// TIA Portal V20 program export: 0 tag tables, 60 data types, 15 data blocks, 199 code blocks (in call order from the OBs), 5 instance data blocks

TYPE "FRK_Access"
// stored: IsFailsafeCompliant false
   STRUCT
      CurrentLevel : DInt;
      CurrentUser : String[32];
      LoginFailed : Bool;
      Policy { S7_SetPoint := 'True'} : "ST_AccessPolicy";
      SessionGeneration : UDInt;
      LoginBusy : Bool;
      LoginResultSequence : UDInt;
      LoginTimeoutMs : UDInt;
      PolicySlot { ExternalAccessible := 'False'; ExternalVisible := 'False'; ExternalWritable := 'False'} : Int;
      PolicyLost { ExternalAccessible := 'False'; ExternalVisible := 'False'; ExternalWritable := 'False'} : Bool;
      PolicyLossAlarm { ExternalAccessible := 'False'; ExternalVisible := 'False'; ExternalWritable := 'False'} : Int;
      UserLossAlarm { ExternalAccessible := 'False'; ExternalVisible := 'False'; ExternalWritable := 'False'} : Int;
      ProviderGeneration { ExternalAccessible := 'False'; ExternalVisible := 'False'; ExternalWritable := 'False'} : UDInt;
      CandidateGeneration { ExternalAccessible := 'False'; ExternalVisible := 'False'; ExternalWritable := 'False'} : UDInt;
      ProviderEnabled { ExternalAccessible := 'False'; ExternalVisible := 'False'; ExternalWritable := 'False'} : Bool;
      LastActivity { ExternalAccessible := 'False'; ExternalVisible := 'False'; ExternalWritable := 'False'} : UDInt;
      LoginSince { ExternalAccessible := 'False'; ExternalVisible := 'False'; ExternalWritable := 'False'} : UDInt;
      LoginSequence { ExternalAccessible := 'False'; ExternalVisible := 'False'; ExternalWritable := 'False'} : UDInt;
      CandidateUser { ExternalAccessible := 'False'; ExternalVisible := 'False'; ExternalWritable := 'False'} : String[32];
      CandidateLevel { ExternalAccessible := 'False'; ExternalVisible := 'False'; ExternalWritable := 'False'} : DInt;
      Round { ExternalAccessible := 'False'; ExternalVisible := 'False'; ExternalWritable := 'False'} : DInt;
      Salt { ExternalAccessible := 'False'; ExternalVisible := 'False'; ExternalWritable := 'False'} : Array[0..15] of Byte;
      Digest { ExternalAccessible := 'False'; ExternalVisible := 'False'; ExternalWritable := 'False'} : Array[0..31] of Byte;
      Expected { ExternalAccessible := 'False'; ExternalVisible := 'False'; ExternalWritable := 'False'} : Array[0..31] of Byte;
   END_STRUCT;
END_TYPE

TYPE "FRK_AccessPolicyImage"
// stored: IsFailsafeCompliant false
   STRUCT
      SchemaVersion { ExternalAccessible := 'False'; ExternalVisible := 'False'; ExternalWritable := 'False'} : UInt;
      Initialized { ExternalAccessible := 'False'; ExternalVisible := 'False'; ExternalWritable := 'False'} : Bool;
      Scope { ExternalAccessible := 'False'; ExternalVisible := 'False'; ExternalWritable := 'False'} : String[80];
      Generation { ExternalAccessible := 'False'; ExternalVisible := 'False'; ExternalWritable := 'False'} : UDInt;
      Policy { ExternalAccessible := 'False'; ExternalVisible := 'False'; ExternalWritable := 'False'; S7_SetPoint := 'True'} : "ST_AccessPolicy";
      Checksum { ExternalAccessible := 'False'; ExternalVisible := 'False'; ExternalWritable := 'False'} : DWord;
   END_STRUCT;
END_TYPE

TYPE "FRK_AlarmLog"
// stored: IsFailsafeCompliant false
   STRUCT
      Active { S7_SetPoint := 'True'} : Array[1..16] of "ST_AlarmEvent";
      NActive : Int;
      Ring { S7_SetPoint := 'True'} : Array[1..64] of "ST_AlarmEvent";
      RingHead : Int;
      Blocking : Bool;
      Truncated : Bool;
      ComeMs { ExternalAccessible := 'False'; ExternalVisible := 'False'; ExternalWritable := 'False'} : Array[1..16] of UDInt;
      Automatic { ExternalAccessible := 'False'; ExternalVisible := 'False'; ExternalWritable := 'False'} : Array[1..16] of Bool;
      Touched { ExternalAccessible := 'False'; ExternalVisible := 'False'; ExternalWritable := 'False'} : Array[1..16] of Bool;
      RingUsed { ExternalAccessible := 'False'; ExternalVisible := 'False'; ExternalWritable := 'False'} : Int;
   END_STRUCT;
END_TYPE

TYPE "FRK_Carrier"
// stored: IsFailsafeCompliant false
   STRUCT
      Enabled { ExternalAccessible := 'False'; ExternalVisible := 'False'; ExternalWritable := 'False'} : Bool;
      Kind { ExternalAccessible := 'False'; ExternalVisible := 'False'; ExternalWritable := 'False'} : DInt;
      Serial { ExternalAccessible := 'False'; ExternalVisible := 'False'; ExternalWritable := 'False'} : UDInt;
      Context { ExternalAccessible := 'False'; ExternalVisible := 'False'; ExternalWritable := 'False'; S7_SetPoint := 'True'} : "ST_PartContext";
      Written { ExternalAccessible := 'False'; ExternalVisible := 'False'; ExternalWritable := 'False'; S7_SetPoint := 'True'} : "ST_PartContext";
      Writes { ExternalAccessible := 'False'; ExternalVisible := 'False'; ExternalWritable := 'False'} : UDInt;
   END_STRUCT;
END_TYPE

TYPE "FRK_ConfigCursor"
// stored: IsFailsafeCompliant false
   STRUCT
      Position { ExternalAccessible := 'False'; ExternalVisible := 'False'; ExternalWritable := 'False'} : DInt;
      First { ExternalAccessible := 'False'; ExternalVisible := 'False'; ExternalWritable := 'False'} : DInt;
   END_STRUCT;
END_TYPE

TYPE "FRK_ConfigSlot"
// stored: IsFailsafeCompliant false
   STRUCT
      SchemaVersion { ExternalAccessible := 'False'; ExternalVisible := 'False'; ExternalWritable := 'False'} : UInt;
      Used { ExternalAccessible := 'False'; ExternalVisible := 'False'; ExternalWritable := 'False'} : Bool;
      ModelCode { ExternalAccessible := 'False'; ExternalVisible := 'False'; ExternalWritable := 'False'} : String[64];
      Record { ExternalAccessible := 'False'; ExternalVisible := 'False'; ExternalWritable := 'False'; S7_SetPoint := 'True'} : "ST_ConfigRecord";
   END_STRUCT;
END_TYPE

TYPE "FRK_ConfigValue"
// stored: IsFailsafeCompliant false
   STRUCT
      Number { ExternalAccessible := 'False'; ExternalVisible := 'False'; ExternalWritable := 'False'} : LInt;
      Flag { ExternalAccessible := 'False'; ExternalVisible := 'False'; ExternalWritable := 'False'} : Bool;
      Text { ExternalAccessible := 'False'; ExternalVisible := 'False'; ExternalWritable := 'False'} : String[80];
   END_STRUCT;
END_TYPE

TYPE "FRK_Core"
// stored: IsFailsafeCompliant false
   STRUCT
      Named { ExternalAccessible := 'False'; ExternalVisible := 'False'; ExternalWritable := 'False'} : Bool;
      Initialized { ExternalAccessible := 'False'; ExternalVisible := 'False'; ExternalWritable := 'False'} : Bool;
      RegIndex { ExternalAccessible := 'False'; ExternalVisible := 'False'; ExternalWritable := 'False'} : DInt;
      ParentIndex { ExternalAccessible := 'False'; ExternalVisible := 'False'; ExternalWritable := 'False'} : DInt;
      ModuleType { ExternalAccessible := 'False'; ExternalVisible := 'False'; ExternalWritable := 'False'} : DInt;
      Exec { ExternalAccessible := 'False'; ExternalVisible := 'False'; ExternalWritable := 'False'} : DInt;
      ExecPrev { ExternalAccessible := 'False'; ExternalVisible := 'False'; ExternalWritable := 'False'} : Bool;
      AbortPrev { ExternalAccessible := 'False'; ExternalVisible := 'False'; ExternalWritable := 'False'} : Bool;
      Armed { ExternalAccessible := 'False'; ExternalVisible := 'False'; ExternalWritable := 'False'} : Bool;
      Command { ExternalAccessible := 'False'; ExternalVisible := 'False'; ExternalWritable := 'False'} : DInt;
      CommandLabel { ExternalAccessible := 'False'; ExternalVisible := 'False'; ExternalWritable := 'False'} : String[120];
      Dispatch { ExternalAccessible := 'False'; ExternalVisible := 'False'; ExternalWritable := 'False'} : Bool;
      EvInit { ExternalAccessible := 'False'; ExternalVisible := 'False'; ExternalWritable := 'False'} : Bool;
      EvCommandStart { ExternalAccessible := 'False'; ExternalVisible := 'False'; ExternalWritable := 'False'} : Bool;
      ReleasePending { ExternalAccessible := 'False'; ExternalVisible := 'False'; ExternalWritable := 'False'} : Bool;
      EvAbort { ExternalAccessible := 'False'; ExternalVisible := 'False'; ExternalWritable := 'False'} : Bool;
      EvAbortInError { ExternalAccessible := 'False'; ExternalVisible := 'False'; ExternalWritable := 'False'} : Bool;
      EvModeExit { ExternalAccessible := 'False'; ExternalVisible := 'False'; ExternalWritable := 'False'} : Bool;
      EvModeChanged { ExternalAccessible := 'False'; ExternalVisible := 'False'; ExternalWritable := 'False'} : Bool;
      "Step" { ExternalAccessible := 'False'; ExternalVisible := 'False'; ExternalWritable := 'False'} : DInt;
      HookResult { ExternalAccessible := 'False'; ExternalVisible := 'False'; ExternalWritable := 'False'} : DInt;
      Held { ExternalAccessible := 'False'; ExternalVisible := 'False'; ExternalWritable := 'False'} : Bool;
      HoldReq { ExternalAccessible := 'False'; ExternalVisible := 'False'; ExternalWritable := 'False'} : Bool;
      HoldReason { ExternalAccessible := 'False'; ExternalVisible := 'False'; ExternalWritable := 'False'} : DInt;
      DiagTouched { ExternalAccessible := 'False'; ExternalVisible := 'False'; ExternalWritable := 'False'} : Bool;
      TimingOpen { ExternalAccessible := 'False'; ExternalVisible := 'False'; ExternalWritable := 'False'} : Bool;
      StartMs { ExternalAccessible := 'False'; ExternalVisible := 'False'; ExternalWritable := 'False'} : UDInt;
      LastNowMs { ExternalAccessible := 'False'; ExternalVisible := 'False'; ExternalWritable := 'False'} : UDInt;
      DeltaMs { ExternalAccessible := 'False'; ExternalVisible := 'False'; ExternalWritable := 'False'} : UDInt;
      ActiveMs { ExternalAccessible := 'False'; ExternalVisible := 'False'; ExternalWritable := 'False'} : UDInt;
      TimeoutMs { ExternalAccessible := 'False'; ExternalVisible := 'False'; ExternalWritable := 'False'} : UDInt;
      Timing { ExternalAccessible := 'False'; ExternalVisible := 'False'; ExternalWritable := 'False'; S7_SetPoint := 'True'} : "ST_ModuleTiming";
      FaultSlot { ExternalAccessible := 'False'; ExternalVisible := 'False'; ExternalWritable := 'False'} : Int;
      FaultHandled { ExternalAccessible := 'False'; ExternalVisible := 'False'; ExternalWritable := 'False'} : Bool;
   END_STRUCT;
END_TYPE

TYPE "FRK_DecisionSlot"
// stored: IsFailsafeCompliant false
   STRUCT
      RootIndex { ExternalAccessible := 'False'; ExternalVisible := 'False'; ExternalWritable := 'False'} : DInt;
      Owner { ExternalAccessible := 'False'; ExternalVisible := 'False'; ExternalWritable := 'False'} : DInt;
      Request { ExternalAccessible := 'False'; ExternalVisible := 'False'; ExternalWritable := 'False'; S7_SetPoint := 'True'} : "ST_DecisionRequest";
      Answer { ExternalAccessible := 'False'; ExternalVisible := 'False'; ExternalWritable := 'False'} : Int;
      AskedAt { ExternalAccessible := 'False'; ExternalVisible := 'False'; ExternalWritable := 'False'} : UDInt;
      OverlapLogged { ExternalAccessible := 'False'; ExternalVisible := 'False'; ExternalWritable := 'False'} : Bool;
      ResolutionLogged { ExternalAccessible := 'False'; ExternalVisible := 'False'; ExternalWritable := 'False'} : Bool;
   END_STRUCT;
END_TYPE

TYPE "FRK_JsonField"
// stored: IsFailsafeCompliant false
   STRUCT
      Key { ExternalAccessible := 'False'; ExternalVisible := 'False'; ExternalWritable := 'False'} : String[16];
      Text { ExternalAccessible := 'False'; ExternalVisible := 'False'; ExternalWritable := 'False'} : WString[160];
      Quoted { ExternalAccessible := 'False'; ExternalVisible := 'False'; ExternalWritable := 'False'} : Bool;
   END_STRUCT;
END_TYPE

TYPE "FRK_ManualConditionRow"
// stored: IsFailsafeCompliant false
   STRUCT
      Used { ExternalAccessible := 'False'; ExternalVisible := 'False'; ExternalWritable := 'False'} : Bool;
      Value { ExternalAccessible := 'False'; ExternalVisible := 'False'; ExternalWritable := 'False'} : DInt;
      Ok { ExternalAccessible := 'False'; ExternalVisible := 'False'; ExternalWritable := 'False'} : Bool;
      Diag { ExternalAccessible := 'False'; ExternalVisible := 'False'; ExternalWritable := 'False'; S7_SetPoint := 'True'} : "ST_Diagnostic";
      Bypassable { ExternalAccessible := 'False'; ExternalVisible := 'False'; ExternalWritable := 'False'} : Bool;
   END_STRUCT;
END_TYPE

TYPE "FRK_PermCtx"
// stored: IsFailsafeCompliant false
   STRUCT
      Permit : Bool;
      Count : Int;
      Blocker : String[160];
   END_STRUCT;
END_TYPE

TYPE "FRK_RegistryRow"
// stored: IsFailsafeCompliant false
   STRUCT
      Valid { ExternalAccessible := 'False'; ExternalVisible := 'False'; ExternalWritable := 'False'} : Bool;
      Parent { ExternalAccessible := 'False'; ExternalVisible := 'False'; ExternalWritable := 'False'} : DInt;
      ModuleType { ExternalAccessible := 'False'; ExternalVisible := 'False'; ExternalWritable := 'False'} : DInt;
      TypeId { ExternalAccessible := 'False'; ExternalVisible := 'False'; ExternalWritable := 'False'} : DInt;
      Capabilities { ExternalAccessible := 'False'; ExternalVisible := 'False'; ExternalWritable := 'False'} : DWord;
      Exec { ExternalAccessible := 'False'; ExternalVisible := 'False'; ExternalWritable := 'False'} : DInt;
      ReasonCode { ExternalAccessible := 'False'; ExternalVisible := 'False'; ExternalWritable := 'False'} : DInt;
      Severity { ExternalAccessible := 'False'; ExternalVisible := 'False'; ExternalWritable := 'False'} : DInt;
      AlarmBlocking { ExternalAccessible := 'False'; ExternalVisible := 'False'; ExternalWritable := 'False'} : Bool;
   END_STRUCT;
END_TYPE

TYPE "FRK_SequenceCtx"
// stored: IsFailsafeCompliant false
   STRUCT
      RunPrevious { ExternalAccessible := 'False'; ExternalVisible := 'False'; ExternalWritable := 'False'} : Bool;
      Running : Bool;
      Restart { ExternalAccessible := 'False'; ExternalVisible := 'False'; ExternalWritable := 'False'} : Bool;
      Done : Bool;
      Error : Bool;
      Pending : Bool;
      StartLatched { ExternalAccessible := 'False'; ExternalVisible := 'False'; ExternalWritable := 'False'} : Bool;
      OwnerIndex { ExternalAccessible := 'False'; ExternalVisible := 'False'; ExternalWritable := 'False'} : DInt;
      ChainIndex { ExternalAccessible := 'False'; ExternalVisible := 'False'; ExternalWritable := 'False'} : DInt;
      "Step" : DInt;
      ScanStep { ExternalAccessible := 'False'; ExternalVisible := 'False'; ExternalWritable := 'False'} : DInt;
      RecordedStep { ExternalAccessible := 'False'; ExternalVisible := 'False'; ExternalWritable := 'False'} : DInt;
      RetVal { ExternalAccessible := 'False'; ExternalVisible := 'False'; ExternalWritable := 'False'} : DInt;
      Scan { ExternalAccessible := 'False'; ExternalVisible := 'False'; ExternalWritable := 'False'} : UDInt;
      Visit { ExternalAccessible := 'False'; ExternalVisible := 'False'; ExternalWritable := 'False'} : UDInt;
      Elapsed : Time;
      DelayElapsed { ExternalAccessible := 'False'; ExternalVisible := 'False'; ExternalWritable := 'False'} : Time;
      StepName : String[160];
      Awaiting : String[160];
      ErrorDiagnostic { S7_SetPoint := 'True'} : "ST_Diagnostic";
      BranchIndex { ExternalAccessible := 'False'; ExternalVisible := 'False'; ExternalWritable := 'False'} : DInt;
      CommandFailed { ExternalAccessible := 'False'; ExternalVisible := 'False'; ExternalWritable := 'False'} : Bool;
      CommandIssued { ExternalAccessible := 'False'; ExternalVisible := 'False'; ExternalWritable := 'False'} : Bool;
      Warned { ExternalAccessible := 'False'; ExternalVisible := 'False'; ExternalWritable := 'False'} : Bool;
      HandledDiagnostic { ExternalAccessible := 'False'; ExternalVisible := 'False'; ExternalWritable := 'False'; S7_SetPoint := 'True'} : "ST_Diagnostic";
      EventVisit { ExternalAccessible := 'False'; ExternalVisible := 'False'; ExternalWritable := 'False'} : UDInt;
      EventToken { ExternalAccessible := 'False'; ExternalVisible := 'False'; ExternalWritable := 'False'} : DInt;
   END_STRUCT;
END_TYPE

TYPE "FRK_SequenceRow"
// stored: IsFailsafeCompliant false
   STRUCT
      StepNo : DInt;
      Visited : Bool;
      LastDuration : Time;
   END_STRUCT;
END_TYPE

TYPE "FRK_SetPayload"
// stored: IsFailsafeCompliant false
   STRUCT
      Info { ExternalAccessible := 'False'; ExternalVisible := 'False'; ExternalWritable := 'False'; S7_SetPoint := 'True'} : "ST_ConfigSetInfo";
      Records { ExternalAccessible := 'False'; ExternalVisible := 'False'; ExternalWritable := 'False'; S7_SetPoint := 'True'} : Array[1..3] of "ST_ConfigRecord";
   END_STRUCT;
END_TYPE

TYPE "FRK_SetWorkspace"
// stored: IsFailsafeCompliant false
   STRUCT
      Payload { ExternalAccessible := 'False'; ExternalVisible := 'False'; ExternalWritable := 'False'; S7_SetPoint := 'True'} : "FRK_SetPayload";
      Seen { ExternalAccessible := 'False'; ExternalVisible := 'False'; ExternalWritable := 'False'} : Array[1..3] of Bool;
      Matched { ExternalAccessible := 'False'; ExternalVisible := 'False'; ExternalWritable := 'False'} : Int;
      RejectScope { ExternalAccessible := 'False'; ExternalVisible := 'False'; ExternalWritable := 'False'} : String[80];
      RejectKey { ExternalAccessible := 'False'; ExternalVisible := 'False'; ExternalWritable := 'False'} : String[160];
      Importing { ExternalAccessible := 'False'; ExternalVisible := 'False'; ExternalWritable := 'False'} : Bool;
      Exporting { ExternalAccessible := 'False'; ExternalVisible := 'False'; ExternalWritable := 'False'} : Bool;
      NextLine { ExternalAccessible := 'False'; ExternalVisible := 'False'; ExternalWritable := 'False'} : Int;
      Generation { ExternalAccessible := 'False'; ExternalVisible := 'False'; ExternalWritable := 'False'} : UDInt;
      Received { ExternalAccessible := 'False'; ExternalVisible := 'False'; ExternalWritable := 'False'} : Int;
      Piece { ExternalAccessible := 'False'; ExternalVisible := 'False'; ExternalWritable := 'False'} : WString[480];
      Line { ExternalAccessible := 'False'; ExternalVisible := 'False'; ExternalWritable := 'False'} : WString[480];
      Fields { ExternalAccessible := 'False'; ExternalVisible := 'False'; ExternalWritable := 'False'; S7_SetPoint := 'True'} : Array[1..9] of "FRK_JsonField";
      FieldCount { ExternalAccessible := 'False'; ExternalVisible := 'False'; ExternalWritable := 'False'} : Int;
   END_STRUCT;
END_TYPE

TYPE "FRK_Unit"
// stored: IsFailsafeCompliant false
   STRUCT
      Initialized { ExternalAccessible := 'False'; ExternalVisible := 'False'; ExternalWritable := 'False'} : Bool;
      Mode { ExternalAccessible := 'False'; ExternalVisible := 'False'; ExternalWritable := 'False'} : DInt;
      RequestedMode { ExternalAccessible := 'False'; ExternalVisible := 'False'; ExternalWritable := 'False'} : DInt;
      ModePending { ExternalAccessible := 'False'; ExternalVisible := 'False'; ExternalWritable := 'False'} : Bool;
      ExitFirst { ExternalAccessible := 'False'; ExternalVisible := 'False'; ExternalWritable := 'False'} : Bool;
      RunReq { ExternalAccessible := 'False'; ExternalVisible := 'False'; ExternalWritable := 'False'} : Bool;
      AbortReq { ExternalAccessible := 'False'; ExternalVisible := 'False'; ExternalWritable := 'False'} : Bool;
      StopReq { ExternalAccessible := 'False'; ExternalVisible := 'False'; ExternalWritable := 'False'} : Bool;
      ModeSince { ExternalAccessible := 'False'; ExternalVisible := 'False'; ExternalWritable := 'False'} : UDInt;
      ReleaseChildren { ExternalAccessible := 'False'; ExternalVisible := 'False'; ExternalWritable := 'False'} : Bool;
      Clearing { ExternalAccessible := 'False'; ExternalVisible := 'False'; ExternalWritable := 'False'} : Bool;
      FaultLatched { ExternalAccessible := 'False'; ExternalVisible := 'False'; ExternalWritable := 'False'} : Bool;
      PrevError { ExternalAccessible := 'False'; ExternalVisible := 'False'; ExternalWritable := 'False'} : Bool;
      EvReset { ExternalAccessible := 'False'; ExternalVisible := 'False'; ExternalWritable := 'False'} : Bool;
      SeenSequence { ExternalAccessible := 'False'; ExternalVisible := 'False'; ExternalWritable := 'False'} : UDInt;
      RequestPending { ExternalAccessible := 'False'; ExternalVisible := 'False'; ExternalWritable := 'False'} : Bool;
      Request { ExternalAccessible := 'False'; ExternalVisible := 'False'; ExternalWritable := 'False'; S7_SetPoint := 'True'} : "ST_HmiRequest";
      RequestUser { ExternalAccessible := 'False'; ExternalVisible := 'False'; ExternalWritable := 'False'} : String[32];
      Permit { ExternalAccessible := 'False'; ExternalVisible := 'False'; ExternalWritable := 'False'} : Bool;
      PermitDiag { ExternalAccessible := 'False'; ExternalVisible := 'False'; ExternalWritable := 'False'; S7_SetPoint := 'True'} : "ST_Diagnostic";
      CarrierIndex { ExternalAccessible := 'False'; ExternalVisible := 'False'; ExternalWritable := 'False'} : DInt;
      Good { ExternalAccessible := 'False'; ExternalVisible := 'False'; ExternalWritable := 'False'} : UDInt;
      Nok { ExternalAccessible := 'False'; ExternalVisible := 'False'; ExternalWritable := 'False'} : UDInt;
      Rework { ExternalAccessible := 'False'; ExternalVisible := 'False'; ExternalWritable := 'False'} : UDInt;
      NokReason { ExternalAccessible := 'False'; ExternalVisible := 'False'; ExternalWritable := 'False'} : DInt;
      CascadePending { ExternalAccessible := 'False'; ExternalVisible := 'False'; ExternalWritable := 'False'} : Bool;
      CascadeKind { ExternalAccessible := 'False'; ExternalVisible := 'False'; ExternalWritable := 'False'} : DInt;
      CascadeMode { ExternalAccessible := 'False'; ExternalVisible := 'False'; ExternalWritable := 'False'} : DInt;
      FollowStart { ExternalAccessible := 'False'; ExternalVisible := 'False'; ExternalWritable := 'False'} : Bool;
      AlarmBlocking { ExternalAccessible := 'False'; ExternalVisible := 'False'; ExternalWritable := 'False'} : Bool;
      ConfigBlocked { ExternalAccessible := 'False'; ExternalVisible := 'False'; ExternalWritable := 'False'} : Bool;
      ConfigEnabled { ExternalAccessible := 'False'; ExternalVisible := 'False'; ExternalWritable := 'False'} : Bool;
      ModelEnabled { ExternalAccessible := 'False'; ExternalVisible := 'False'; ExternalWritable := 'False'} : Bool;
      ConfigSetsEnabled { ExternalAccessible := 'False'; ExternalVisible := 'False'; ExternalWritable := 'False'} : Bool;
   END_STRUCT;
END_TYPE

TYPE "ST_AccessPolicy"
// stored: IsFailsafeCompliant false
   STRUCT
      Required : Array[0..11] of DInt;
      SessionTimeout : Time := T#0MS;
   END_STRUCT;
END_TYPE

TYPE "ST_AlarmEvent"
// stored: IsFailsafeCompliant false
   STRUCT
      ReasonCode : DInt;
      Description : WString[255];
      SourcePath : WString[255];
      IoTag : String[80];
      IoAddress : String[80];
      Severity : DInt;
      Category : DInt;
      ResetClass : DInt;
      State : DInt;
      ComeAt : LDT;
      GoneAt : LDT;
      ResetAt : LDT;
      Duration : Time;
      Shelved : Bool;
      ShelvedUntil : LDT;
      ComeTimeSynchronized : Bool;
      GoneTimeSynchronized : Bool;
      ResetTimeSynchronized : Bool;
      ShelfTimeSynchronized : Bool;
   END_STRUCT;
END_TYPE

TYPE "ST_CommandInfo"
// stored: IsFailsafeCompliant false
   STRUCT
      Value : DInt;
      Label : String[120];
      Style : DInt;
   END_STRUCT;
END_TYPE

TYPE "ST_ConfigEntry"
// stored: IsFailsafeCompliant false
   STRUCT
      Scope : WString[255];
      Item : WString[255];
      ValueText : WString[255];
      WriteKey : String[160];
      WriteRevision : UDInt;
      ConfigKind : DInt;
      ValueType : DInt;
      Writable : Bool;
      RequiresReady : Bool;
      HasMinimum : Bool;
      HasMaximum : Bool;
      Minimum : LReal;
      Maximum : LReal;
      Unit : String[16];
      LabelKey : String[160];
      EnumDomain : WString[255];
      ClassId : String[40];
      ReadLevel : DInt;
      WriteLevel : DInt;
      Readable : Bool;
      UnitCode : DInt;
      EnumLabelKey : String[80];
      ModelScoped : Bool;
   END_STRUCT;
END_TYPE

TYPE "ST_ConfigPage"
// stored: IsFailsafeCompliant false
   STRUCT
      Revision : UDInt;
      PageIndex : Int;
      PageCount : Int;
      EntryCount : Int;
      Entries { S7_SetPoint := 'True'} : Array[1..16] of "ST_ConfigEntry";
   END_STRUCT;
END_TYPE

TYPE "ST_ConfigPersistStatus"
// stored: IsFailsafeCompliant false
   STRUCT
      Pending : Bool;
      Failed : Bool;
      WindowMs : UDInt := 5000;
      PendingSince : LDT;
      StorePresent : Bool;
      StoreKind : DInt;
      RestorePolicy : DInt;
      RestoreLost : Bool;
      RestoreAcknowledged : Bool;
      LostPath : String[80];
      LastSetName : String[80];
      LastSetRecords : Int;
      LastRejectScope : String[80];
      LastRejectKey : String[160];
   END_STRUCT;
END_TYPE

TYPE "ST_ConfigRecord"
// stored: IsFailsafeCompliant false
   STRUCT
      Scope : String[80];
      WriteKey : String[160];
      Revision : UDInt;
      Kind : DInt;
      ValueType : DInt;
      ValueText : String[80];
   END_STRUCT;
END_TYPE

TYPE "ST_ConfigSetInfo"
// stored: IsFailsafeCompliant false
   STRUCT
      Used : Bool;
      SetName : String[80];
      RootIdentity : String[80];
      SetSchema : UInt;
      ConfigRev : UDInt;
      Kind : DInt;
      ModelCode : String[64];
      RecordCount : Int;
      CreatedAt : LDT;
      TimeSynchronized : Bool;
   END_STRUCT;
END_TYPE

TYPE "ST_CylinderDevice"
// stored: IsFailsafeCompliant false
   STRUCT
      Direction : DInt;
      Withdrawn : Bool;
      Extended : Bool;
      Retracted : Bool;
      Lease { S7_SetPoint := 'True'} : "ST_SequenceCommandLease";
   END_STRUCT;
END_TYPE

TYPE "ST_CylinderHal"
// stored: IsFailsafeCompliant false
   STRUCT
      FeedbackExtended : Bool;
      FeedbackRetracted : Bool;
      ExtendPermit : Bool;
      RetractPermit : Bool;
      PermitDiagnostic { S7_SetPoint := 'True'} : "ST_Diagnostic";
      RetractDiagnostic { S7_SetPoint := 'True'} : "ST_Diagnostic";
      CoilExtend : Bool;
      CoilRetract : Bool;
   END_STRUCT;
END_TYPE

TYPE "ST_CylinderOutCmd"
// stored: IsFailsafeCompliant false
   STRUCT
      Direction : DInt;
   END_STRUCT;
END_TYPE

TYPE "ST_CylinderOutImm"
// stored: IsFailsafeCompliant false
   STRUCT
      Extended : Bool;
      Retracted : Bool;
   END_STRUCT;
END_TYPE

TYPE "ST_CylinderParCfg"
// stored: IsFailsafeCompliant false
   STRUCT
      SchemaVersion : UInt := 1;
      Timeout : Time := T#8S;
   END_STRUCT;
END_TYPE

TYPE "ST_CylinderParCmd"
// stored: IsFailsafeCompliant false
   STRUCT
      Reserved : Bool;
   END_STRUCT;
END_TYPE

TYPE "ST_DecisionRequest"
// stored: IsFailsafeCompliant false
   STRUCT
      Prompt : WString[255];
      Options : Array[1..6] of String[64];
      Default : Int;
      Timeout : Time;
      SourcePath : WString[255];
   END_STRUCT;
END_TYPE

TYPE "ST_Diagnostic"
// stored: IsFailsafeCompliant false
   STRUCT
      ReasonCode : DInt;
      SourcePath : WString[255];
      Description : WString[255];
      IoTag : String[80];
      IoAddress : String[80];
      Severity : DInt;
      Category : DInt;
      Since : LDT;
      TimeSynchronized : Bool;
   END_STRUCT;
END_TYPE

TYPE "ST_FraktalHal"
// stored: IsFailsafeCompliant false
   STRUCT
      PressDemo { ExternalAccessible := 'False'; ExternalVisible := 'False'; ExternalWritable := 'False'; S7_SetPoint := 'True'} : "ST_PressDemoUnitHal";
   END_STRUCT;
END_TYPE

TYPE "ST_HmiRequest"
// stored: IsFailsafeCompliant false
   STRUCT
      Kind : DInt;
      TargetPath : WString[255];
      NameValue : String[160];
      TextValue : WString[255];
      User : String[32];
      Secret : String[32];
      IntValue : DInt;
      BoolValue : Bool;
      DurationMs : UDInt;
      Sequence : UDInt;
   END_STRUCT;
END_TYPE

TYPE "ST_HmiResponse"
// stored: IsFailsafeCompliant false
   STRUCT
      AckSequence : UDInt;
      Accepted : Bool;
      Diagnostic : WString[255];
      Report { S7_SetPoint := 'True'} : "ST_ReleaseReport";
      ConfigPage { S7_SetPoint := 'True'} : "ST_ConfigPage";
   END_STRUCT;
END_TYPE

TYPE "ST_MeasRecord"
// stored: IsFailsafeCompliant false
   STRUCT
      "Name" : String[64];
      Value : LReal;
      Minimum : LReal;
      Maximum : LReal;
      Target : LReal;
      Unit : String[16];
      InTol : Bool;
   END_STRUCT;
END_TYPE

TYPE "ST_ModePolicy"
// stored: IsFailsafeCompliant false
   STRUCT
      Shield : DInt;
      Style : DInt;
   END_STRUCT;
END_TYPE

TYPE "ST_ModelField"
// stored: IsFailsafeCompliant false
   STRUCT
      "Name" : String[32];
      Value : String[64];
   END_STRUCT;
END_TYPE

TYPE "ST_ModelId"
// stored: IsFailsafeCompliant false
   STRUCT
      ModelCode : String[64];
      "Family" : String[64];
      Variant : String[64];
      Fields { S7_SetPoint := 'True'} : Array[1..8] of "ST_ModelField";
      NField : Int;
   END_STRUCT;
END_TYPE

TYPE "ST_ModuleStatus"
// stored: IsFailsafeCompliant false
   STRUCT
      "Name" : String[80];
      DisplayNameKey : String[160];
      DescriptionKey : String[160];
      TypeKey : String[160];
      ModuleType : DInt;
      State : DInt;
      FaultActive : Bool;
      Diagnostic { S7_SetPoint := 'True'} : "ST_Diagnostic";
      TileEnable : Bool := TRUE;
      ControlDomainId : String[80];
   END_STRUCT;
END_TYPE

TYPE "ST_ModuleTiming"
// stored: IsFailsafeCompliant false
   STRUCT
      LastCmdTime : Time;
      Rows { S7_SetPoint := 'True'} : Array[1..8] of "ST_TimingRow";
      Truncated : Bool;
   END_STRUCT;
END_TYPE

TYPE "ST_PartContext"
// stored: IsFailsafeCompliant false
   STRUCT
      Uid : String[64];
      Present : Bool;
      CarrierKind : DInt;
      Result { S7_SetPoint := 'True'} : "ST_PartResult";
      Parents : Array[1..8] of String[64];
   END_STRUCT;
END_TYPE

TYPE "ST_PartResult"
// stored: IsFailsafeCompliant false
   STRUCT
      Verdict : DInt;
      ReasonCode : DInt;
      Records { S7_SetPoint := 'True'} : Array[1..32] of "ST_MeasRecord";
      StationPath : WString[255];
      Stamp : LDT;
      TimeSynchronized : Bool;
   END_STRUCT;
END_TYPE

TYPE "ST_PressDemoCycle"
// stored: IsFailsafeCompliant false
   STRUCT
      PartInMachine { ExternalAccessible := 'False'; ExternalVisible := 'False'; ExternalWritable := 'False'} : Bool;
      PartDispositioned { ExternalAccessible := 'False'; ExternalVisible := 'False'; ExternalWritable := 'False'} : Bool;
      CycleCompleted { ExternalAccessible := 'False'; ExternalVisible := 'False'; ExternalWritable := 'False'} : Bool;
      FailureReason { ExternalAccessible := 'False'; ExternalVisible := 'False'; ExternalWritable := 'False'} : DInt;
   END_STRUCT;
END_TYPE

TYPE "ST_PressDemoOutCmd"
// stored: IsFailsafeCompliant false
   STRUCT
      CycleCompleted : Bool;
   END_STRUCT;
END_TYPE

TYPE "ST_PressDemoOutImm"
// stored: IsFailsafeCompliant false
   STRUCT
      Homed : Bool;
   END_STRUCT;
END_TYPE

TYPE "ST_PressDemoParCfg"
// stored: IsFailsafeCompliant false
   STRUCT
      SchemaVersion : UInt := 1;
      Timeout : Time := T#0MS;
   END_STRUCT;
END_TYPE

TYPE "ST_PressDemoParCmd"
// stored: IsFailsafeCompliant false
   STRUCT
      Reserved : Bool;
   END_STRUCT;
END_TYPE

TYPE "ST_PressDemoReleaseConditions"
// stored: IsFailsafeCompliant false
   STRUCT
      ModeStartAirPressureOk : Bool;
      RamGuardClosed : Bool;
      RamSlideInside : Bool;
      RamDevicesHealthy : Bool;
      RamAirPressureOk : Bool;
      RamTwoHandHeld : Bool;
   END_STRUCT;
END_TYPE

TYPE "ST_PressDemoSignals"
// stored: IsFailsafeCompliant false
   STRUCT
      PartPresent { ExternalAccessible := 'False'; ExternalVisible := 'False'; ExternalWritable := 'False'} : Bool;
      PartQuality { ExternalAccessible := 'False'; ExternalVisible := 'False'; ExternalWritable := 'False'} : Bool;
      AirPressureOk { ExternalAccessible := 'False'; ExternalVisible := 'False'; ExternalWritable := 'False'} : Bool;
      TwoHandHeld { ExternalAccessible := 'False'; ExternalVisible := 'False'; ExternalWritable := 'False'} : Bool;
      StartPulse { ExternalAccessible := 'False'; ExternalVisible := 'False'; ExternalWritable := 'False'} : Bool;
      PermitDiagnostic { ExternalAccessible := 'False'; ExternalVisible := 'False'; ExternalWritable := 'False'; S7_SetPoint := 'True'} : "ST_Diagnostic";
   END_STRUCT;
END_TYPE

TYPE "ST_PressDemoStationCfg"
// stored: IsFailsafeCompliant false
   STRUCT
      SchemaVersion : UInt := 1;
      RequireTwoHandStart : Bool := TRUE;
      TransferSettleTime : Time := T#200MS;
      PressSettleTime : Time := T#300MS;
   END_STRUCT;
END_TYPE

TYPE "ST_PressDemoUnitHal"
// stored: IsFailsafeCompliant false
   STRUCT
      PressRam { ExternalAccessible := 'False'; ExternalVisible := 'False'; ExternalWritable := 'False'; S7_SetPoint := 'True'} : "ST_CylinderHal";
      Door { ExternalAccessible := 'False'; ExternalVisible := 'False'; ExternalWritable := 'False'; S7_SetPoint := 'True'} : "ST_CylinderHal";
      PartSlide { ExternalAccessible := 'False'; ExternalVisible := 'False'; ExternalWritable := 'False'; S7_SetPoint := 'True'} : "ST_CylinderHal";
      Process { ExternalAccessible := 'False'; ExternalVisible := 'False'; ExternalWritable := 'False'; S7_SetPoint := 'True'} : "ST_PressDemoSignals";
   END_STRUCT;
END_TYPE

TYPE "ST_ReleaseReason"
// stored: IsFailsafeCompliant false
   STRUCT
      Description : WString[255];
      ReasonCode : DInt;
      SourcePath : WString[255];
      Kind : DInt;
      Bypassable : Bool;
   END_STRUCT;
END_TYPE

TYPE "ST_ReleaseReport"
// stored: IsFailsafeCompliant false
   STRUCT
      Released : Bool;
      Count : Int;
      Reasons { S7_SetPoint := 'True'} : Array[1..24] of "ST_ReleaseReason";
   END_STRUCT;
END_TYPE

TYPE "ST_SequenceCommandLease"
// stored: IsFailsafeCompliant false
   STRUCT
      OwnerIndex : DInt;
      ChainIndex : DInt;
      BranchIndex : DInt;
      "Step" : DInt;
      Raised : Bool;
      AbortIssued : Bool;
      ReleasedScan : UDInt;
   END_STRUCT;
END_TYPE

TYPE "ST_StateFlag"
// stored: IsFailsafeCompliant false
   STRUCT
      Key : String[120];
      Value : Bool;
      Since : LDT;
      Stale : Bool;
   END_STRUCT;
END_TYPE

TYPE "ST_TimingRow"
// stored: IsFailsafeCompliant false
   STRUCT
      Id : DInt;
      Label : String[120];
      TimeClass : DInt;
      Count : UDInt;
      Last : Time;
      Minimum : Time;
      Maximum : Time;
      Avg : Time;
   END_STRUCT;
END_TYPE

TYPE "ST_UserRecord"
// stored: IsFailsafeCompliant false
   STRUCT
      User : String[32];
      Salt : Array[0..15] of Byte;
      PinHash : Array[0..31] of Byte;
      Level : DInt;
   END_STRUCT;
END_TYPE

DATA_BLOCK "FRK_AccessPolicies"   // DB3
{ S7_Optimized_Access := 'TRUE' }
VERSION : 0.1
// stored: AutoNumber true, DBAccessibleFromOPCUA true, DBAccessibleFromWebserver true, IsOnlyStoredInLoadMemory false, IsRetainMemResEnabled false, IsWriteProtectedInAS false, MemoryReserve 100
   VAR RETAIN
      Rows { ExternalAccessible := 'False'; ExternalVisible := 'False'; ExternalWritable := 'False'; S7_SetPoint := 'True'} : Array[1..1] of "FRK_AccessPolicyImage";
   END_VAR
BEGIN
END_DATA_BLOCK

DATA_BLOCK "FRK_AccessStorage"   // DB4
{ S7_Optimized_Access := 'TRUE' }
VERSION : 0.1
// stored: AutoNumber true, DBAccessibleFromOPCUA true, DBAccessibleFromWebserver true, IsOnlyStoredInLoadMemory false, IsRetainMemResEnabled false, IsWriteProtectedInAS false, MemoryReserve 100
   VAR
      UsersReady { ExternalAccessible := 'False'; ExternalVisible := 'False'; ExternalWritable := 'False'} : Bool;
      UsersLost { ExternalAccessible := 'False'; ExternalVisible := 'False'; ExternalWritable := 'False'} : Bool;
      EmptyPolicy { ExternalAccessible := 'False'; ExternalVisible := 'False'; ExternalWritable := 'False'; S7_SetPoint := 'True'} : "ST_AccessPolicy";
   END_VAR
   VAR RETAIN
      UsersCommissioned { ExternalAccessible := 'False'; ExternalVisible := 'False'; ExternalWritable := 'False'} : Bool;
   END_VAR
BEGIN
END_DATA_BLOCK

DATA_BLOCK "FRK_Carriers"   // DB5
{ S7_Optimized_Access := 'TRUE' }
VERSION : 0.1
// stored: AutoNumber true, DBAccessibleFromOPCUA true, DBAccessibleFromWebserver true, IsOnlyStoredInLoadMemory false, IsRetainMemResEnabled false, IsWriteProtectedInAS false, MemoryReserve 100
   VAR
      Slots { ExternalAccessible := 'False'; ExternalVisible := 'False'; ExternalWritable := 'False'; S7_SetPoint := 'True'} : Array[0..4] of "FRK_Carrier";
   END_VAR
BEGIN
END_DATA_BLOCK

DATA_BLOCK "FRK_Clock"   // DB1
{ S7_Optimized_Access := 'TRUE' }
VERSION : 0.1
// stored: AutoNumber true, DBAccessibleFromOPCUA true, DBAccessibleFromWebserver true, IsOnlyStoredInLoadMemory false, IsRetainMemResEnabled false, IsWriteProtectedInAS false, MemoryReserve 100
   VAR
      Mem { ExternalAccessible := 'False'; ExternalVisible := 'False'; ExternalWritable := 'False'} : LReal;
      AccMs { ExternalAccessible := 'False'; ExternalVisible := 'False'; ExternalWritable := 'False'} : LReal;
      NowMs { ExternalAccessible := 'False'; ExternalVisible := 'False'; ExternalWritable := 'False'} : UDInt;
   END_VAR
BEGIN
END_DATA_BLOCK

DATA_BLOCK "FRK_ConfigRuntime"   // DB6
{ S7_Optimized_Access := 'TRUE' }
VERSION : 0.1
// stored: AutoNumber true, DBAccessibleFromOPCUA true, DBAccessibleFromWebserver true, IsOnlyStoredInLoadMemory false, IsRetainMemResEnabled false, IsWriteProtectedInAS false, MemoryReserve 100
   VAR
      Fresh { ExternalAccessible := 'False'; ExternalVisible := 'False'; ExternalWritable := 'False'} : Bool;
      Unavailable { ExternalAccessible := 'False'; ExternalVisible := 'False'; ExternalWritable := 'False'} : Bool;
      Failed { ExternalAccessible := 'False'; ExternalVisible := 'False'; ExternalWritable := 'False'} : Array[1..1] of Bool;
      LossSlot { ExternalAccessible := 'False'; ExternalVisible := 'False'; ExternalWritable := 'False'} : Array[1..1] of Int;
   END_VAR
BEGIN
END_DATA_BLOCK

DATA_BLOCK "FRK_ConfigScratch"   // DB7
{ S7_Optimized_Access := 'TRUE' }
VERSION : 0.1
// stored: AutoNumber true, DBAccessibleFromOPCUA true, DBAccessibleFromWebserver true, IsOnlyStoredInLoadMemory false, IsRetainMemResEnabled false, IsWriteProtectedInAS false, MemoryReserve 100
   VAR
      Entry { ExternalAccessible := 'False'; ExternalVisible := 'False'; ExternalWritable := 'False'; S7_SetPoint := 'True'} : "ST_ConfigEntry";
      Blank { ExternalAccessible := 'False'; ExternalVisible := 'False'; ExternalWritable := 'False'; S7_SetPoint := 'True'} : "ST_ConfigEntry";
      Value { ExternalAccessible := 'False'; ExternalVisible := 'False'; ExternalWritable := 'False'; S7_SetPoint := 'True'} : "FRK_ConfigValue";
      Storage { ExternalAccessible := 'False'; ExternalVisible := 'False'; ExternalWritable := 'False'} : DInt;
      Schema { ExternalAccessible := 'False'; ExternalVisible := 'False'; ExternalWritable := 'False'} : UInt;
      Minimum { ExternalAccessible := 'False'; ExternalVisible := 'False'; ExternalWritable := 'False'} : LReal;
      Maximum { ExternalAccessible := 'False'; ExternalVisible := 'False'; ExternalWritable := 'False'} : LReal;
      MaxLength { ExternalAccessible := 'False'; ExternalVisible := 'False'; ExternalWritable := 'False'} : Int;
      MinRead { ExternalAccessible := 'False'; ExternalVisible := 'False'; ExternalWritable := 'False'} : DInt;
      MinWrite { ExternalAccessible := 'False'; ExternalVisible := 'False'; ExternalWritable := 'False'} : DInt;
   END_VAR
BEGIN
END_DATA_BLOCK

DATA_BLOCK "FRK_ConfigStore"   // DB8
{ S7_Optimized_Access := 'TRUE' }
VERSION : 0.1
// stored: AutoNumber true, DBAccessibleFromOPCUA true, DBAccessibleFromWebserver true, IsOnlyStoredInLoadMemory false, IsRetainMemResEnabled false, IsWriteProtectedInAS false, MemoryReserve 100
   VAR RETAIN
      SchemaVersion { ExternalAccessible := 'False'; ExternalVisible := 'False'; ExternalWritable := 'False'} : UInt;
      Rows { ExternalAccessible := 'False'; ExternalVisible := 'False'; ExternalWritable := 'False'; S7_SetPoint := 'True'} : Array[1..3] of "FRK_ConfigSlot";
      ActiveModels { ExternalAccessible := 'False'; ExternalVisible := 'False'; ExternalWritable := 'False'} : Array[1..1] of String[64];
      Lost { ExternalAccessible := 'False'; ExternalVisible := 'False'; ExternalWritable := 'False'} : Array[1..1] of Bool;
      Acknowledged { ExternalAccessible := 'False'; ExternalVisible := 'False'; ExternalWritable := 'False'} : Array[1..1] of Bool;
      LostPath { ExternalAccessible := 'False'; ExternalVisible := 'False'; ExternalWritable := 'False'} : Array[1..1] of String[80];
   END_VAR
BEGIN
END_DATA_BLOCK

DATA_BLOCK "FRK_Decisions"   // DB9
{ S7_Optimized_Access := 'TRUE' }
VERSION : 0.1
// stored: AutoNumber true, DBAccessibleFromOPCUA true, DBAccessibleFromWebserver true, IsOnlyStoredInLoadMemory false, IsRetainMemResEnabled false, IsWriteProtectedInAS false, MemoryReserve 100
   VAR
      Slots { ExternalAccessible := 'False'; ExternalVisible := 'False'; ExternalWritable := 'False'; S7_SetPoint := 'True'} : Array[1..1] of "FRK_DecisionSlot";
      EmptyRequest { ExternalAccessible := 'False'; ExternalVisible := 'False'; ExternalWritable := 'False'; S7_SetPoint := 'True'} : "ST_DecisionRequest";
   END_VAR
BEGIN
END_DATA_BLOCK

DATA_BLOCK "FRK_LocalUsers"   // DB10
{ S7_Optimized_Access := 'TRUE' }
VERSION : 0.1
// stored: AutoNumber true, DBAccessibleFromOPCUA true, DBAccessibleFromWebserver true, IsOnlyStoredInLoadMemory false, IsRetainMemResEnabled false, IsWriteProtectedInAS false, MemoryReserve 100
   VAR RETAIN
      SchemaVersion { ExternalAccessible := 'False'; ExternalVisible := 'False'; ExternalWritable := 'False'} : UInt;
      Generation { ExternalAccessible := 'False'; ExternalVisible := 'False'; ExternalWritable := 'False'} : UDInt;
      Count { ExternalAccessible := 'False'; ExternalVisible := 'False'; ExternalWritable := 'False'} : DInt;
      Rows { ExternalAccessible := 'False'; ExternalVisible := 'False'; ExternalWritable := 'False'; S7_SetPoint := 'True'} : Array[1..16] of "ST_UserRecord";
      Checksum { ExternalAccessible := 'False'; ExternalVisible := 'False'; ExternalWritable := 'False'} : DWord;
   END_VAR
BEGIN
END_DATA_BLOCK

DATA_BLOCK "FRK_Registry"   // DB2
{ S7_Optimized_Access := 'TRUE' }
VERSION : 0.1
// stored: AutoNumber true, DBAccessibleFromOPCUA true, DBAccessibleFromWebserver true, IsOnlyStoredInLoadMemory false, IsRetainMemResEnabled false, IsWriteProtectedInAS false, MemoryReserve 100
   VAR
      Count { ExternalAccessible := 'False'; ExternalVisible := 'False'; ExternalWritable := 'False'} : DInt;
      Fault { ExternalAccessible := 'False'; ExternalVisible := 'False'; ExternalWritable := 'False'} : Bool;
      Rows { ExternalAccessible := 'False'; ExternalVisible := 'False'; ExternalWritable := 'False'; S7_SetPoint := 'True'} : Array[0..4] of "FRK_RegistryRow";
   END_VAR
BEGIN
END_DATA_BLOCK

DATA_BLOCK "FRK_SetRuntime"   // DB11
{ S7_Optimized_Access := 'TRUE' }
VERSION : 0.1
// stored: AutoNumber true, DBAccessibleFromOPCUA true, DBAccessibleFromWebserver true, IsOnlyStoredInLoadMemory false, IsRetainMemResEnabled false, IsWriteProtectedInAS false, MemoryReserve 100
   VAR
      Work { ExternalAccessible := 'False'; ExternalVisible := 'False'; ExternalWritable := 'False'; S7_SetPoint := 'True'} : Array[1..1] of "FRK_SetWorkspace";
   END_VAR
BEGIN
END_DATA_BLOCK

DATA_BLOCK "FRK_SetStore"   // DB12
{ S7_Optimized_Access := 'TRUE' }
VERSION : 0.1
// stored: AutoNumber true, DBAccessibleFromOPCUA true, DBAccessibleFromWebserver true, IsOnlyStoredInLoadMemory false, IsRetainMemResEnabled false, IsWriteProtectedInAS false, MemoryReserve 100
   VAR RETAIN
      SchemaVersion { ExternalAccessible := 'False'; ExternalVisible := 'False'; ExternalWritable := 'False'} : UInt;
      Sets { ExternalAccessible := 'False'; ExternalVisible := 'False'; ExternalWritable := 'False'; S7_SetPoint := 'True'} : Array[1..1, 1..4] of "FRK_SetPayload";
   END_VAR
BEGIN
END_DATA_BLOCK

DATA_BLOCK "FRK_UnitScratch"   // DB13
{ S7_Optimized_Access := 'TRUE' }
VERSION : 0.1
// stored: AutoNumber true, DBAccessibleFromOPCUA true, DBAccessibleFromWebserver true, IsOnlyStoredInLoadMemory false, IsRetainMemResEnabled false, IsWriteProtectedInAS false, MemoryReserve 100
   VAR
      Response { ExternalAccessible := 'False'; ExternalVisible := 'False'; ExternalWritable := 'False'; S7_SetPoint := 'True'} : "ST_HmiResponse";
      EmptyDiagnostic { ExternalAccessible := 'False'; ExternalVisible := 'False'; ExternalWritable := 'False'; S7_SetPoint := 'True'} : "ST_Diagnostic";
      EmptyConfigEntry { ExternalAccessible := 'False'; ExternalVisible := 'False'; ExternalWritable := 'False'; S7_SetPoint := 'True'} : "ST_ConfigEntry";
      EmptyEvent { ExternalAccessible := 'False'; ExternalVisible := 'False'; ExternalWritable := 'False'; S7_SetPoint := 'True'} : "ST_AlarmEvent";
   END_VAR
BEGIN
END_DATA_BLOCK

DATA_BLOCK "GDB_FraktalHal"   // DB16
{ S7_Optimized_Access := 'TRUE' }
VERSION : 0.1
// stored: AutoNumber true, DBAccessibleFromOPCUA true, DBAccessibleFromWebserver true, IsOnlyStoredInLoadMemory false, IsRetainMemResEnabled false, IsWriteProtectedInAS false, MemoryReserve 100
   VAR
      Data { ExternalAccessible := 'False'; ExternalVisible := 'False'; ExternalWritable := 'False'; S7_SetPoint := 'True'} : "ST_FraktalHal";
   END_VAR
BEGIN
END_DATA_BLOCK

DATA_BLOCK "GDB_PressDemoIO"   // DB19
{ S7_Optimized_Access := 'TRUE' }
VERSION : 0.1
// Demo logical I/O boundary. Bind these symbols to the commissioned hardware
//  driver when a bench is available; feedback is never synthesized here.
// stored: AutoNumber true, DBAccessibleFromOPCUA true, DBAccessibleFromWebserver true, IsOnlyStoredInLoadMemory false, IsRetainMemResEnabled false, IsWriteProtectedInAS false, MemoryReserve 100
   VAR
      PartPresent : Bool;
      PartQuality : Bool;
      AirPressureOk : Bool;
      TwoHandHeld : Bool;
      StartPulse : Bool;
      RamExtended : Bool;
      RamRetracted : Bool;
      DoorClosed : Bool;
      DoorOpen : Bool;
      SlideInside : Bool;
      SlideOutside : Bool;
      RamExtend : Bool;
      RamRetract : Bool;
      DoorClose : Bool;
      DoorRelease : Bool;
      SlideExtend : Bool;
      SlideRetract : Bool;
   END_VAR
BEGIN
END_DATA_BLOCK

ORGANIZATION_BLOCK "Main"   // OB1, SCL, ProgramCycle
TITLE = "Main Program Sweep (Cycle)"
{ S7_Optimized_Access := 'TRUE' }
VERSION : 0.1
// stored: AutoNumber true, IsIECCheckEnabled false, SetENOAutomatically false
   VAR_INPUT
      Initial_Call : Bool;   // Initial call of this OB
      Remanence : Bool;   // =True, if remanent data are available
   END_VAR
BEGIN

   "F_PressDemoReadInputs"();
   "GDB_FraktalMain"(Startup := #Initial_Call);
   "F_PressDemoWriteOutputs"();
END_ORGANIZATION_BLOCK

FUNCTION_BLOCK "FB_FraktalMain"   // FB13, SCL
{ S7_Optimized_Access := 'TRUE' }
VERSION : 0.1
// stored: AutoNumber true, IsIECCheckEnabled false, IsRetainMemResEnabled false, MemoryReserve 100, SetENOAutomatically false, UDAEnableTagReadback false
   VAR_INPUT
      Startup { ExternalAccessible := 'False'; ExternalVisible := 'False'; ExternalWritable := 'False'} : Bool;
   END_VAR
BEGIN

   IF #Startup THEN
       "FRK_Registry".Count := 0;
       "FRK_Registry".Fault := FALSE;
   END_IF;
   "FRK_ClockTick"();
   "FRK_AccessStoreBoot"(Startup := #Startup);
   "FRK_ConfigBoot"(Startup := #Startup);
   "FRK_SetBoot"(Startup := #Startup);
   "PressDemo"(ParentIndex := 0,
               Startup := #Startup,
               Hal := "GDB_FraktalHal".Data.PressDemo);
END_FUNCTION_BLOCK

FUNCTION_BLOCK "FB_PressDemoUnit"   // FB12, SCL
{ S7_Optimized_Access := 'TRUE' }
VERSION : 0.1
// Generated frame v0.11; change the declaration, then regenerate.
// stored: AutoNumber true, IsIECCheckEnabled false, IsRetainMemResEnabled false, MemoryReserve 100, SetENOAutomatically false, UDAEnableTagReadback false
   VAR_INPUT
      Execute { ExternalWritable := 'False'} : Bool;
      Abort { ExternalWritable := 'False'} : Bool;
      Command { ExternalWritable := 'False'} : DInt;
      ParCfg { ExternalWritable := 'False'} : "ST_PressDemoParCfg";
      ParCmd { ExternalWritable := 'False'} : "ST_PressDemoParCmd";
      ParentIndex { ExternalAccessible := 'False'; ExternalVisible := 'False'; ExternalWritable := 'False'} : DInt;
      Startup { ExternalAccessible := 'False'; ExternalVisible := 'False'; ExternalWritable := 'False'} : Bool;
   END_VAR
   VAR_OUTPUT
      Busy { ExternalWritable := 'False'} : Bool;
      Done { ExternalWritable := 'False'} : Bool;
      Error { ExternalWritable := 'False'} : Bool;
      Aborted { ExternalWritable := 'False'} : Bool;
      Held { ExternalWritable := 'False'} : Bool;
      ErrorID { ExternalWritable := 'False'} : DWord;
      Timing { ExternalWritable := 'False'} : "ST_ModuleTiming";
      OutCmd { ExternalWritable := 'False'} : "ST_PressDemoOutCmd";
      OutImm { ExternalWritable := 'False'} : "ST_PressDemoOutImm";
   END_VAR
   VAR_IN_OUT
      Hal : "ST_PressDemoUnitHal";
   END_VAR
   VAR
      Status { ExternalWritable := 'False'; S7_SetPoint := 'True'} : "ST_ModuleStatus";
      Core { ExternalAccessible := 'False'; ExternalVisible := 'False'; ExternalWritable := 'False'; S7_SetPoint := 'True'} : "FRK_Core";
      LatchedParCmd { ExternalAccessible := 'False'; ExternalVisible := 'False'; ExternalWritable := 'False'; S7_SetPoint := 'True'} : "ST_PressDemoParCmd";
      StateFlags { ExternalWritable := 'False'; S7_SetPoint := 'True'} : Array[1..12] of "ST_StateFlag";
      StateFlagCount { ExternalWritable := 'False'} : Int;
      StateTouched { ExternalAccessible := 'False'; ExternalVisible := 'False'; ExternalWritable := 'False'} : Array[1..12] of Bool;
      StationCfg { ExternalWritable := 'False'; S7_SetPoint := 'True'} : "ST_PressDemoStationCfg";
      ConfigStageStationCfg { ExternalAccessible := 'False'; ExternalVisible := 'False'; ExternalWritable := 'False'; S7_SetPoint := 'True'} : "ST_PressDemoStationCfg";
      ConfigDefaultStationCfg { ExternalAccessible := 'False'; ExternalVisible := 'False'; ExternalWritable := 'False'; S7_SetPoint := 'True'} : "ST_PressDemoStationCfg";
      ConfigStaged { ExternalAccessible := 'False'; ExternalVisible := 'False'; ExternalWritable := 'False'} : Bool;
      ConfigPersist { ExternalWritable := 'False'; S7_SetPoint := 'True'} : "ST_ConfigPersistStatus";
      ModelId { ExternalWritable := 'False'; S7_SetPoint := 'True'} : "ST_ModelId";
      AvailableModelCount { ExternalWritable := 'False'} : Int;
      AvailableModels { ExternalWritable := 'False'; S7_SetPoint := 'True'} : Array[1..1] of "ST_ModelId";
      ConfigSets { ExternalWritable := 'False'; S7_SetPoint := 'True'} : Array[1..4] of "ST_ConfigSetInfo";
      ConfigSetCount { ExternalWritable := 'False'} : Int;
      ConfigSetDocument { ExternalWritable := 'False'} : WString[480];
      ConfigSetDocumentLine { ExternalWritable := 'False'} : Int;
      ConfigSetDocumentLines { ExternalWritable := 'False'} : Int;
      Unit { ExternalAccessible := 'False'; ExternalVisible := 'False'; ExternalWritable := 'False'; S7_SetPoint := 'True'} : "FRK_Unit";
      Auto { ExternalWritable := 'False'; S7_SetPoint := 'True'} : "FB_PressDemoAutoGraphOwner";
      Home { ExternalWritable := 'False'; S7_SetPoint := 'True'} : "FB_PressDemoHomeGraphOwner";
      Release { ExternalWritable := 'False'; S7_SetPoint := 'True'} : "FB_PressDemoRelease";
      SequenceReset { ExternalAccessible := 'False'; ExternalVisible := 'False'; ExternalWritable := 'False'} : Bool;
      HmiRequest { S7_SetPoint := 'True'} : "ST_HmiRequest";
      ModePolicy { ExternalAccessible := 'False'; ExternalVisible := 'False'; ExternalWritable := 'False'; S7_SetPoint := 'True'} : Array[0..6] of "ST_ModePolicy";
      Access { ExternalWritable := 'False'; S7_SetPoint := 'True'} : "FRK_Access";
      HmiResponse { ExternalWritable := 'False'; S7_SetPoint := 'True'} : "ST_HmiResponse";
      ConfigRev { ExternalWritable := 'False'} : UDInt;
      ConfigCursor { ExternalAccessible := 'False'; ExternalVisible := 'False'; ExternalWritable := 'False'; S7_SetPoint := 'True'} : "FRK_ConfigCursor";
      Part { ExternalWritable := 'False'; S7_SetPoint := 'True'} : "ST_PartContext";
      Decision { ExternalWritable := 'False'; S7_SetPoint := 'True'} : "ST_DecisionRequest";
      DecisionAnswer { ExternalWritable := 'False'} : Int;
      History { ExternalWritable := 'False'; S7_SetPoint := 'True'} : Array[1..16] of "ST_Diagnostic";
      HistoryHead { ExternalWritable := 'False'} : Int;
      AlarmLog { ExternalWritable := 'False'; S7_SetPoint := 'True'} : "FRK_AlarmLog";
      ModeActivePublished { ExternalWritable := 'False'} : DInt;
      RunningPublished { ExternalWritable := 'False'} : Bool;
      StopPendingPublished { ExternalWritable := 'False'} : Bool;
      SupportedModesPublished { ExternalWritable := 'False'} : Array[0..6] of Bool;
      GoodCount { ExternalWritable := 'False'} : UDInt;
      NokCount { ExternalWritable := 'False'} : UDInt;
      ReworkCount { ExternalWritable := 'False'} : UDInt;
      NokReason { ExternalWritable := 'False'} : DInt;
      PressRam { ExternalWritable := 'False'; S7_SetPoint := 'True'} : "FB_CylinderCM";
      Door { ExternalWritable := 'False'; S7_SetPoint := 'True'} : "FB_CylinderCM";
      PartSlide { ExternalWritable := 'False'; S7_SetPoint := 'True'} : "FB_CylinderCM";
   END_VAR
   VAR_TEMP
      InstancePath : WString[254];
      RouteMatched : Bool;
      ManualMatched : Bool;
      ConfigRootIndex : Int;
   END_VAR
   VAR CONSTANT
      EXEC_READY : DInt := 0;
      MODULE_TIER : DInt := 1;
   END_VAR
BEGIN

   // ---- GENERATED: setup
   IF #Startup OR NOT #Core.Named THEN
       #InstancePath := GetInstancePath(size := 0);
       "FRK_SetIdentity"(Core := #Core,
                         Status := #Status,
                         InstancePath := #InstancePath,
                         ModuleType := 1,
                         TypeId := 1,
                         Capabilities := DWORD#16#00000000,
                         ParentIndex := #ParentIndex,
                         TypeKey := 'project.pressDemo');
   END_IF;
   IF #Startup THEN "FRK_CfgRestore_PressDemoUnit"(Core := #Core,
                                                       Status := #Status,
                                                       StationCfg := #StationCfg,
                                                       ConfigStageStationCfg := #ConfigStageStationCfg,
                                                       ConfigDefaultStationCfg := #ConfigDefaultStationCfg);
   END_IF;
   #ConfigRootIndex := "FRK_ConfigRoot"(RegIndex := #Core.RegIndex);
   IF #Core.ParentIndex = 0 THEN
       #AvailableModelCount := 0;
   ELSE
       #AvailableModelCount := 0;
   END_IF;
   "FRK_StateSweep"(Flags := #StateFlags,
                    Count := #StateFlagCount,
                    Touched := #StateTouched,
                    Startup := #Startup);
   IF #Startup OR #ConfigRev = 0 THEN
       #ConfigRev := "FRK_ConfigRevision"(Previous := #ConfigRev);
   END_IF;
   #SupportedModesPublished[0] := TRUE;
   #SupportedModesPublished[1] := TRUE;
   #SupportedModesPublished[2] := TRUE;
   #SupportedModesPublished[3] := FALSE;
   #SupportedModesPublished[4] := FALSE;
   #SupportedModesPublished[5] := FALSE;
   #SupportedModesPublished[6] := FALSE;
   "FRK_UnitPrepare"(Core := #Core,
                     Unit := #Unit,
                     Policy := #ModePolicy,
                     Request := #HmiRequest,
                     Response := #HmiResponse,
                     Startup := #Startup,
                     InitialMode := 1);
   "FRK_AlarmBegin"(AlarmLog := #AlarmLog,
                    Startup := #Startup);
   "FRK_AccessPolicyBoot"(Access := #Access,
                          Startup := #Startup,
                          Root := #Core.ParentIndex = 0,
                          Scope := #Status.Name);
   "FRK_AccessCyclic"(Access := #Access,
                      Startup := #Startup,
                      SourcePath := STRING_TO_WSTRING(#Status.Name),
                      AlarmLog := #AlarmLog,
                      Revision := #ConfigRev);
   "FRK_UnitMailbox"(Core := #Core,
                     Unit := #Unit,
                     Status := #Status,
                     Policy := #ModePolicy,
                     Access := #Access,
                     Request := #HmiRequest,
                     Response := #HmiResponse,
                     Supported := #SupportedModesPublished);
   "FRK_ConfigStatus"(RootIndex := #ConfigRootIndex,
                      Scope := #Status.Name,
                      PolicyLost := #Access.PolicyLost,
                      UsersLost := "FRK_AccessStorage".UsersLost,
                      Persist := #ConfigPersist,
                      AlarmLog := #AlarmLog);
   #Unit.ConfigEnabled := #Core.ParentIndex = 0;
   #Unit.ConfigSetsEnabled := TRUE AND #Core.ParentIndex = 0;
   #Unit.ModelEnabled := #AvailableModelCount > 0;
   #Unit.ConfigBlocked := #ConfigPersist.RestoreLost AND NOT #ConfigPersist.RestoreAcknowledged AND #ConfigPersist.RestorePolicy = 1;
   #Unit.ConfigBlocked := #Unit.ConfigBlocked OR #Access.PolicyLost;
   // ---- GENERATED: begin
   "FRK_Begin"(Core := #Core,
               Status := #Status,
               Execute := #Unit.RunReq,
               Abort := (#Abort OR #Unit.AbortReq),
               Command := 1);
   IF #Core.EvCommandStart THEN
       #LatchedParCmd := #ParCmd;
       CASE #Core.Command OF
           1:
               "FRK_UnitRunStart"(Core := #Core,
                                  Status := #Status,
                                  Timeout := #ParCfg.Timeout,
                                  Label := 'Run');
           ELSE
               "FRK_Start"(Core := #Core,
                           Status := #Status,
                           Supported := FALSE,
                           Timeout := T#0ms,
                           Label := '');
       END_CASE;
   END_IF;
   // ---- AUTHORED: cyclic management
   #Release(AirPressureOk := #Hal.Process.AirPressureOk,
            DoorClosed := #Hal.Door.FeedbackExtended AND NOT #Hal.Door.FeedbackRetracted,
            SlideInside := #Hal.PartSlide.FeedbackExtended AND NOT #Hal.PartSlide.FeedbackRetracted,
            RamHealthy := NOT #PressRam.Error AND NOT #PressRam.Aborted,
            DoorHealthy := NOT #Door.Error AND NOT #Door.Aborted,
            SlideHealthy := NOT #PartSlide.Error AND NOT #PartSlide.Aborted,
            TwoHandHeld := #Hal.Process.TwoHandHeld OR NOT #StationCfg.RequireTwoHandStart);
   #Hal.Process.PermitDiagnostic := "FRK_UnitScratch".EmptyDiagnostic;
   #Hal.Process.PermitDiagnostic.Description := STRING_TO_WSTRING(#Release.ModeStart.Blocker);
   #Hal.Process.PermitDiagnostic.SourcePath := STRING_TO_WSTRING(#Status.Name);
   #Hal.PressRam.ExtendPermit := #Release.RamExtend.Permit;
   #Hal.PressRam.RetractPermit := #Hal.Process.AirPressureOk;
   #Hal.PressRam.PermitDiagnostic := "FRK_UnitScratch".EmptyDiagnostic;
   #Hal.PressRam.PermitDiagnostic.Description := STRING_TO_WSTRING(#Release.RamExtend.Blocker);
   #Hal.PressRam.PermitDiagnostic.SourcePath := STRING_TO_WSTRING(#Status.Name);
   #Hal.PressRam.RetractDiagnostic := #Hal.Process.PermitDiagnostic;
   #Hal.Door.PermitDiagnostic := #Hal.Process.PermitDiagnostic;
   #Hal.Door.RetractDiagnostic := #Hal.Process.PermitDiagnostic;
   #Hal.PartSlide.PermitDiagnostic := #Hal.Process.PermitDiagnostic;
   #Hal.PartSlide.RetractDiagnostic := #Hal.Process.PermitDiagnostic;
   #Hal.Door.ExtendPermit := #Hal.Process.AirPressureOk;
   #Hal.Door.RetractPermit := #Hal.Process.AirPressureOk;
   #Hal.PartSlide.ExtendPermit := #Hal.Process.AirPressureOk;
   #Hal.PartSlide.RetractPermit := #Hal.Process.AirPressureOk;
   // ---- GENERATED: end management
   "FRK_Release_PressDemoUnit"(Unit := #Unit,
                               Hal := #Hal);
   IF #Core.RegIndex > 0 THEN
       "FRK_Registry".Rows[#Core.RegIndex].AlarmBlocking := #AlarmLog.Blocking;
   END_IF;
   #Unit.AlarmBlocking := "FRK_AlarmTreeBlocking"(Owner := #Core.RegIndex);
   "FRK_UnitConsume"(Core := #Core,
                     Unit := #Unit,
                     Status := #Status,
                     Policy := #ModePolicy,
                     Access := #Access,
                     Response := #HmiResponse,
                     Supported := #SupportedModesPublished);
   "FRK_UnitMode"(Core := #Core,
                  Unit := #Unit);
   "FRK_UnitModeResolve"(Core := #Core,
                         Unit := #Unit,
                         Status := #Status,
                         Policy := #ModePolicy,
                         Timeout := #ParCfg.Timeout);
   "FRK_DecisionCyclic"(Owner := #Core.RegIndex,
                        Busy := #Core.Exec = 1,
                        Reset := #Startup OR #Unit.EvReset OR #Core.EvModeChanged,
                        AlarmLog := #AlarmLog);
   "FRK_UnitFollow"(Core := #Core,
                    Unit := #Unit,
                    Status := #Status,
                    Policy := #ModePolicy,
                    Access := #Access,
                    Supported := #SupportedModesPublished);
   IF #Unit.RequestPending AND (#Unit.Request.Kind = 11 OR #Unit.Request.Kind = 16) THEN
       #ManualMatched := FALSE;
       #RouteMatched := "FRK_Route_CylinderCM"(Module := #PressRam, Hal := #Hal.PressRam, Request := #Unit.Request, Report := #HmiResponse.Report);
       #ManualMatched := #ManualMatched OR #RouteMatched;
       #RouteMatched := "FRK_Route_CylinderCM"(Module := #Door, Hal := #Hal.Door, Request := #Unit.Request, Report := #HmiResponse.Report);
       #ManualMatched := #ManualMatched OR #RouteMatched;
       #RouteMatched := "FRK_Route_CylinderCM"(Module := #PartSlide, Hal := #Hal.PartSlide, Request := #Unit.Request, Report := #HmiResponse.Report);
       #ManualMatched := #ManualMatched OR #RouteMatched;
       IF NOT #ManualMatched THEN
           "FRK_ReleaseReason"(Report := #HmiResponse.Report,
                               Description := WSTRING#'std.error.unsupportedHmiRequest',
                               Reason := 2008,
                               Path := #Unit.Request.TargetPath,
                               Kind := 4);
       END_IF;
       #HmiResponse.Accepted := #Unit.Request.Kind = 16 OR #HmiResponse.Report.Released;
       IF #Unit.Request.Kind = 11 THEN
           IF #HmiResponse.Accepted THEN
               #HmiResponse.Diagnostic := WSTRING#'std.audit.manualCommandAccepted';
           ELSE
               #HmiResponse.Diagnostic := WSTRING#'std.audit.manualCommandRejected';
           END_IF;
       END_IF;
   END_IF;
   IF #Unit.EvReset THEN
       "FRK_AlarmOperatorReset"(AlarmLog := #AlarmLog);
   END_IF;
   IF #Core.ReleasePending OR #Unit.ReleaseChildren THEN
       "FRK_ReleaseCommand"(Core := #PressRam.Core,
                            Execute := #PressRam.Execute);
       "FRK_ReleaseCommand"(Core := #Door.Core,
                            Execute := #Door.Execute);
       "FRK_ReleaseCommand"(Core := #PartSlide.Core,
                            Execute := #PartSlide.Execute);
   END_IF;
   // ---- GENERATED: child call
   #PressRam(ParentIndex := #Core.RegIndex,
             Startup := #Startup,
             Hal := #Hal.PressRam);
   "FRK_ManualFinish"(Core := #PressRam.Core,
                      Execute := #PressRam.Execute,
                      ManualOwned := #PressRam.ManualOwned);
   // ---- GENERATED: child call
   #Door(ParentIndex := #Core.RegIndex,
         Startup := #Startup,
         Hal := #Hal.Door);
   "FRK_ManualFinish"(Core := #Door.Core,
                      Execute := #Door.Execute,
                      ManualOwned := #Door.ManualOwned);
   // ---- GENERATED: child call
   #PartSlide(ParentIndex := #Core.RegIndex,
              Startup := #Startup,
              Hal := #Hal.PartSlide);
   "FRK_ManualFinish"(Core := #PartSlide.Core,
                      Execute := #PartSlide.Execute,
                      ManualOwned := #PartSlide.ManualOwned);
   #Unit.CascadePending := FALSE;
   "FRK_CfgOperation_PressDemoUnit"(Core := #Core, Status := #Status, ModePolicy := #ModePolicy, Access := #Access, Unit := #Unit, HmiResponse := #HmiResponse, ConfigPersist := #ConfigPersist, ConfigCursor := #ConfigCursor, ConfigRev := #ConfigRev, ModelId := #ModelId, AvailableModelCount := #AvailableModelCount, StationCfg := #StationCfg, PressRam := #PressRam, Door := #Door, PartSlide := #PartSlide);
   "FRK_CfgSetOperation_PressDemoUnit"(Core := #Core, Status := #Status, ModePolicy := #ModePolicy, Access := #Access, Unit := #Unit, HmiResponse := #HmiResponse, ConfigPersist := #ConfigPersist, ConfigRev := #ConfigRev, ModelId := #ModelId, ConfigSets := #ConfigSets, ConfigSetCount := #ConfigSetCount, ConfigSetDocument := #ConfigSetDocument, ConfigSetDocumentLine := #ConfigSetDocumentLine, ConfigSetDocumentLines := #ConfigSetDocumentLines, SupportedModesPublished := #SupportedModesPublished, StationCfg := #StationCfg, ConfigStageStationCfg := #ConfigStageStationCfg, PressRam := #PressRam, Door := #Door, PartSlide := #PartSlide, Startup := #Startup);
   IF #Unit.RequestPending AND #Core.ParentIndex = 0 THEN
       "FRK_SetResult"(Request := #Unit.Request,
                       Response := #HmiResponse,
                       Persist := #ConfigPersist,
                       AlarmLog := #AlarmLog,
                       Scope := #Status.Name,
                       RootIndex := #ConfigRootIndex);
   END_IF;
   "FRK_ConfigStatus"(RootIndex := #ConfigRootIndex,
                      Scope := #Status.Name,
                      PolicyLost := #Access.PolicyLost,
                      UsersLost := "FRK_AccessStorage".UsersLost,
                      Persist := #ConfigPersist,
                      AlarmLog := #AlarmLog);
   "FRK_RouteAbort"(Core := #Core,
                    Abort := (#Abort OR #Unit.AbortReq));
   IF #Core.EvAbort THEN
       "FRK_PartAborted"(Core := #Core,
                         Unit := #Unit,
                         Status := #Status,
                         Part := #Part,
                         AlarmLog := #AlarmLog);
   END_IF;
   // ---- AUTHORED: unconditional sequence policy
   #SequenceReset := #Startup OR #Unit.EvReset OR #Core.EvModeChanged OR #Core.EvCommandStart;
   #Auto(Run := #Core.Exec = 1 AND #Unit.Mode = 0 AND NOT "FRK_Registry".Fault,
         Reset := #SequenceReset,
         OwnerIndex := #Core.RegIndex,
         Delta := DINT_TO_TIME(UDINT_TO_DINT(#Core.DeltaMs)),
         PartPresent := #Hal.Process.PartPresent,
         PartQuality := #Hal.Process.PartQuality,
         AirPressureOk := #Hal.Process.AirPressureOk,
         TwoHandHeld := #Hal.Process.TwoHandHeld,
         StartPulse := #Hal.Process.StartPulse,
         RequireTwoHandStart := #StationCfg.RequireTwoHandStart,
         TransferSettleTime := #StationCfg.TransferSettleTime,
         PressSettleTime := #StationCfg.PressSettleTime,
         SourcePath := #Status.Name,
         PressRam := #PressRam,
         Door := #Door,
         PartSlide := #PartSlide,
         Core := #Core,
         Unit := #Unit,
         Status := #Status,
         Part := #Part,
         AlarmLog := #AlarmLog,
         Chart := "GDB_GRAPH_PressDemoAuto");
   #Home(Run := #Core.Exec = 1 AND #Unit.Mode = 2 AND NOT "FRK_Registry".Fault,
         Reset := #SequenceReset,
         OwnerIndex := #Core.RegIndex,
         Delta := DINT_TO_TIME(UDINT_TO_DINT(#Core.DeltaMs)),
         PressRam := #PressRam,
         Door := #Door,
         PartSlide := #PartSlide,
         Chart := "GDB_GRAPH_PressDemoHome");
   "FRK_SeqOwnerStatus"(Seq := #Home.Seq,
                        Core := #Core,
                        Status := #Status);
   IF #Home.Seq.Done AND #Core.Exec = 1 AND #Unit.Mode = 2 THEN
       "FRK_Complete"(Core := #Core,
                      Status := #Status);
   END_IF;
   #OutCmd.CycleCompleted := #Auto.Cycle.CycleCompleted;
   // ---- GENERATED: sequence policy end
   "FRK_End"(Core := #Core,
             Status := #Status,
             Busy => #Busy,
             Done => #Done,
             Error => #Error,
             Aborted => #Aborted,
             Held => #Held,
             ErrorID => #ErrorID,
             Timing => #Timing);
   "FRK_DecisionCyclic"(Owner := #Core.RegIndex,
                        Busy := #Core.Exec = 1,
                        Reset := #Startup OR #Unit.EvReset OR #Core.EvModeChanged,
                        AlarmLog := #AlarmLog);
   "FRK_DecisionPublish"(Owner := #Core.RegIndex,
                         Decision := #Decision,
                         DecisionAnswer := #DecisionAnswer);
   IF NOT #Unit.EvReset THEN
       "FRK_AlarmCapture"(AlarmLog := #AlarmLog,
                          Core := #Core,
                          Status := #Status);
       "FRK_Capture_CylinderCM"(Module := #PressRam,
                                AlarmLog := #AlarmLog);
       "FRK_Capture_CylinderCM"(Module := #Door,
                                AlarmLog := #AlarmLog);
       "FRK_Capture_CylinderCM"(Module := #PartSlide,
                                AlarmLog := #AlarmLog);
       "FRK_AlarmEnd"(AlarmLog := #AlarmLog);
   END_IF;
   IF #Core.RegIndex > 0 THEN
       "FRK_Registry".Rows[#Core.RegIndex].AlarmBlocking := #AlarmLog.Blocking;
   END_IF;
   #Unit.AlarmBlocking := "FRK_AlarmTreeBlocking"(Owner := #Core.RegIndex);
   "FRK_AccessPersist"(Access := #Access,
                       Unit := #Unit,
                       Response := #HmiResponse,
                       SourcePath := STRING_TO_WSTRING(#Status.Name),
                       AlarmLog := #AlarmLog);
   "FRK_AccessFinish"(Access := #Access,
                      Unit := #Unit,
                      Response := #HmiResponse,
                      SourcePath := STRING_TO_WSTRING(#Status.Name),
                      AlarmLog := #AlarmLog,
                      Revision := #ConfigRev);
   "FRK_UnitFinish"(Core := #Core,
                    Unit := #Unit,
                    Response := #HmiResponse,
                    Status := #Status,
                    Part := #Part,
                    AlarmLog := #AlarmLog,
                    History := #History,
                    Head := #HistoryHead);
   #ModeActivePublished := #Unit.Mode;
   #RunningPublished := #Core.Exec = 1;
   #StopPendingPublished := #Unit.StopReq AND #Core.Exec = 1;
   #GoodCount := #Unit.Good;
   #NokCount := #Unit.Nok;
   #ReworkCount := #Unit.Rework;
   #NokReason := #Unit.NokReason;
   // ---- AUTHORED: unconditional cyclic/derived data
   #OutImm.Homed := "FRK_State"(Idx := 1, Key := 'project.state.pressAtLoadPosition',
                                Ok := #PressRam.OutImm.Retracted AND #Door.OutImm.Retracted AND #PartSlide.OutImm.Retracted, Flags := #StateFlags, Count := #StateFlagCount, Touched := #StateTouched);
   // ---- GENERATED: frame end
END_FUNCTION_BLOCK

FUNCTION_BLOCK "FB_PressDemoRelease"   // FB5, SCL
{ S7_Optimized_Access := 'TRUE' }
VERSION : 0.1
// stored: AutoNumber true, IsIECCheckEnabled false, IsRetainMemResEnabled false, MemoryReserve 100, SetENOAutomatically false, UDAEnableTagReadback false
   VAR_INPUT
      AirPressureOk : Bool;
      DoorClosed : Bool;
      DoorHealthy : Bool;
      RamHealthy : Bool;
      SlideHealthy : Bool;
      SlideInside : Bool;
      TwoHandHeld : Bool;
   END_VAR
   VAR
      Conditions { ExternalWritable := 'False'; S7_SetPoint := 'True'} : "ST_PressDemoReleaseConditions";
      ModeStart { ExternalWritable := 'False'; S7_SetPoint := 'True'} : "FRK_PermCtx";
      RamExtend { ExternalWritable := 'False'; S7_SetPoint := 'True'} : "FRK_PermCtx";
   END_VAR
BEGIN

   #Conditions.ModeStartAirPressureOk := #AirPressureOk;
   #Conditions.RamGuardClosed := #DoorClosed;
   #Conditions.RamSlideInside := #SlideInside;
   #Conditions.RamDevicesHealthy := #RamHealthy AND #DoorHealthy AND #SlideHealthy;
   #Conditions.RamAirPressureOk := #AirPressureOk;
   #Conditions.RamTwoHandHeld := #TwoHandHeld;
   "FRK_PermBegin"(Perm := #ModeStart);
   "FRK_PermCondition"(Perm := #ModeStart,
                       Label := 'project.condition.ModeStartAirPressureOk',
                       Ok := #Conditions.ModeStartAirPressureOk);
   "FRK_PermBegin"(Perm := #RamExtend);
   "FRK_PermCondition"(Perm := #RamExtend,
                       Label := 'project.condition.RamGuardClosed',
                       Ok := #Conditions.RamGuardClosed);
   "FRK_PermCondition"(Perm := #RamExtend,
                       Label := 'project.condition.RamSlideInside',
                       Ok := #Conditions.RamSlideInside);
   "FRK_PermCondition"(Perm := #RamExtend,
                       Label := 'project.condition.RamDevicesHealthy',
                       Ok := #Conditions.RamDevicesHealthy);
   "FRK_PermCondition"(Perm := #RamExtend,
                       Label := 'project.condition.RamAirPressureOk',
                       Ok := #Conditions.RamAirPressureOk);
   "FRK_PermCondition"(Perm := #RamExtend,
                       Label := 'project.condition.RamTwoHandHeld',
                       Ok := #Conditions.RamTwoHandHeld);
END_FUNCTION_BLOCK

FUNCTION_BLOCK "FB_CylinderCM"   // FB1, SCL
{ S7_Optimized_Access := 'TRUE' }
VERSION : 0.1
// Generated frame v0.11; change the declaration, then regenerate.
// stored: AutoNumber true, IsIECCheckEnabled false, IsRetainMemResEnabled false, MemoryReserve 100, SetENOAutomatically false, UDAEnableTagReadback false
   VAR_INPUT
      Execute { ExternalWritable := 'False'} : Bool;
      Abort { ExternalWritable := 'False'} : Bool;
      Command { ExternalWritable := 'False'} : DInt;
      ParCfg { ExternalWritable := 'False'} : "ST_CylinderParCfg";
      ParCmd { ExternalWritable := 'False'} : "ST_CylinderParCmd";
      ParentIndex { ExternalAccessible := 'False'; ExternalVisible := 'False'; ExternalWritable := 'False'} : DInt;
      Startup { ExternalAccessible := 'False'; ExternalVisible := 'False'; ExternalWritable := 'False'} : Bool;
   END_VAR
   VAR_OUTPUT
      Busy { ExternalWritable := 'False'} : Bool;
      Done { ExternalWritable := 'False'} : Bool;
      Error { ExternalWritable := 'False'} : Bool;
      Aborted { ExternalWritable := 'False'} : Bool;
      Held { ExternalWritable := 'False'} : Bool;
      ErrorID { ExternalWritable := 'False'} : DWord;
      Timing { ExternalWritable := 'False'} : "ST_ModuleTiming";
      OutCmd { ExternalWritable := 'False'} : "ST_CylinderOutCmd";
      OutImm { ExternalWritable := 'False'} : "ST_CylinderOutImm";
   END_VAR
   VAR_IN_OUT
      Hal : "ST_CylinderHal";
   END_VAR
   VAR
      Status { ExternalWritable := 'False'; S7_SetPoint := 'True'} : "ST_ModuleStatus";
      Core { ExternalAccessible := 'False'; ExternalVisible := 'False'; ExternalWritable := 'False'; S7_SetPoint := 'True'} : "FRK_Core";
      LatchedParCmd { ExternalAccessible := 'False'; ExternalVisible := 'False'; ExternalWritable := 'False'; S7_SetPoint := 'True'} : "ST_CylinderParCmd";
      StateFlags { ExternalWritable := 'False'; S7_SetPoint := 'True'} : Array[1..12] of "ST_StateFlag";
      StateFlagCount { ExternalWritable := 'False'} : Int;
      StateTouched { ExternalAccessible := 'False'; ExternalVisible := 'False'; ExternalWritable := 'False'} : Array[1..12] of Bool;
      Device { ExternalAccessible := 'False'; ExternalVisible := 'False'; ExternalWritable := 'False'; S7_SetPoint := 'True'} : "ST_CylinderDevice";
      Catalog { ExternalAccessible := 'False'; ExternalVisible := 'False'; ExternalWritable := 'False'; S7_SetPoint := 'True'} : Array[1..12] of "ST_CommandInfo";
      CatalogCount { ExternalAccessible := 'False'; ExternalVisible := 'False'; ExternalWritable := 'False'} : Int;
      ManConditions { ExternalAccessible := 'False'; ExternalVisible := 'False'; ExternalWritable := 'False'; S7_SetPoint := 'True'} : Array[1..16] of "FRK_ManualConditionRow";
      ManualOwned { ExternalAccessible := 'False'; ExternalVisible := 'False'; ExternalWritable := 'False'} : Bool;
   END_VAR
   VAR_TEMP
      InstancePath : WString[254];
   END_VAR
   VAR CONSTANT
      EXEC_READY : DInt := 0;
      MODULE_TIER : DInt := 3;
   END_VAR
BEGIN

   // ---- GENERATED: setup
   IF #Startup OR NOT #Core.Named THEN
       #InstancePath := GetInstancePath(size := 0);
       "FRK_SetIdentity"(Core := #Core,
                         Status := #Status,
                         InstancePath := #InstancePath,
                         ModuleType := 3,
                         TypeId := 2,
                         Capabilities := DWORD#16#00000000,
                         ParentIndex := #ParentIndex,
                         TypeKey := 'fraktal.module.cylinder');
       #CatalogCount := 2;
       #Catalog[1].Value := 1;
       #Catalog[1].Label := 'EXTEND';
       #Catalog[1].Style := 0;
       #Catalog[2].Value := 2;
       #Catalog[2].Label := 'RETRACT';
       #Catalog[2].Style := 0;
   END_IF;
   "FRK_StateSweep"(Flags := #StateFlags,
                    Count := #StateFlagCount,
                    Touched := #StateTouched,
                    Startup := #Startup);
   // ---- GENERATED: begin
   "FRK_Begin"(Core := #Core,
               Status := #Status,
               Execute := #Execute,
               Abort := #Abort,
               Command := #Command);
   IF #Core.EvCommandStart THEN
       #LatchedParCmd := #ParCmd;
       CASE #Core.Command OF
           1:
               "FRK_Start"(Core := #Core,
                           Status := #Status,
                           Supported := TRUE,
                           Timeout := #ParCfg.Timeout,
                           Label := 'EXTEND');
           2:
               "FRK_Start"(Core := #Core,
                           Status := #Status,
                           Supported := TRUE,
                           Timeout := #ParCfg.Timeout,
                           Label := 'RETRACT');
           ELSE
               "FRK_Start"(Core := #Core,
                           Status := #Status,
                           Supported := FALSE,
                           Timeout := T#0ms,
                           Label := '');
       END_CASE;
   END_IF;
   IF #Core.EvCommandStart THEN
       // ---- AUTHORED: CommandStart
       #Device.Direction := #Core.Command;
       #Device.Withdrawn := FALSE;
       IF NOT #Device.Lease.Raised THEN
           #Device.Lease.OwnerIndex := 0;
           #Device.Lease.ChainIndex := 0;
           #Device.Lease.BranchIndex := 0;
       END_IF;

       // ---- GENERATED: reaction end
   END_IF;
   // ---- AUTHORED: cyclic management
   #Device.Extended := #Hal.FeedbackExtended AND NOT #Hal.FeedbackRetracted;
   #Device.Retracted := #Hal.FeedbackRetracted AND NOT #Hal.FeedbackExtended;

   // ---- GENERATED: end management
   "FRK_RouteAbort"(Core := #Core,
                    Abort := #Abort);
   IF #Core.EvAbort THEN
       // ---- AUTHORED: Abort
       #Device.Direction := 0;

       // ---- GENERATED: reaction end
   END_IF;
   IF #Core.EvAbortInError THEN
       // ---- AUTHORED: AbortInError
       #Device.Direction := 0;

       // ---- GENERATED: reaction end
   END_IF;
   IF #Core.Dispatch AND #Core.RegIndex > 0 AND NOT "FRK_Registry".Fault THEN
       // ---- AUTHORED: dispatch
       CASE #Core.Command OF
           1:
               IF NOT #Hal.ExtendPermit THEN
                   "FRK_HoldDiag"(Core := #Core,
                                  Status := #Status,
                                  Diag := #Hal.PermitDiagnostic);
               ELSIF #Device.Extended THEN
                   #OutCmd.Direction := #Device.Direction;
                   "FRK_Complete"(Core := #Core,
                                  Status := #Status);
               END_IF;
           2:
               IF NOT #Hal.RetractPermit THEN
                   "FRK_HoldDiag"(Core := #Core,
                                  Status := #Status,
                                  Diag := #Hal.RetractDiagnostic);
               ELSIF #Device.Retracted THEN
                   #OutCmd.Direction := #Device.Direction;
                   "FRK_Complete"(Core := #Core,
                                  Status := #Status);
               END_IF;
           ELSE
               // The shared frame rejects unknown commands before dispatch.
               #Device.Direction := 0;
       END_CASE;

       // ---- GENERATED: end dispatch
   END_IF;
   "FRK_End"(Core := #Core,
             Status := #Status,
             Busy => #Busy,
             Done => #Done,
             Error => #Error,
             Aborted => #Aborted,
             Held => #Held,
             ErrorID => #ErrorID,
             Timing => #Timing);
   // ---- AUTHORED: unconditional cyclic/derived data
   // Apply the SAME live permit to latched coils after completion as while BUSY.
   #Hal.CoilExtend := #Device.Direction = 1 AND #Hal.ExtendPermit
   AND NOT #Device.Withdrawn AND #Core.Exec <> 3 AND #Core.Exec <> 4;
   #Hal.CoilRetract := #Device.Direction = 2 AND #Hal.RetractPermit
   AND NOT #Device.Withdrawn AND #Core.Exec <> 3 AND #Core.Exec <> 4;
   #OutImm.Extended := "FRK_State"(Idx := 1, Key := 'module.state.extended',
                                   Ok := #Device.Extended, Flags := #StateFlags, Count := #StateFlagCount, Touched := #StateTouched);
   #OutImm.Retracted := "FRK_State"(Idx := 2, Key := 'module.state.retracted',
                                    Ok := #Device.Retracted, Flags := #StateFlags, Count := #StateFlagCount, Touched := #StateTouched);

   // ---- GENERATED: frame end
END_FUNCTION_BLOCK

FUNCTION_BLOCK "FB_PressDemoAutoGraphOwner"   // FB10, SCL
{ S7_Optimized_Access := 'TRUE' }
VERSION : 0.1
// stored: AutoNumber true, IsIECCheckEnabled false, IsRetainMemResEnabled false, MemoryReserve 100, SetENOAutomatically false, UDAEnableTagReadback false
   VAR_INPUT
      Run : Bool;
      Reset : Bool;
      OwnerIndex : DInt;
      Delta : Time;
      TransferSettleTime : Time;
      PartQuality : Bool;
      RequireTwoHandStart : Bool;
      SourcePath : String[80];
      PartPresent : Bool;
      AirPressureOk : Bool;
      TwoHandHeld : Bool;
      StartPulse : Bool;
      PressSettleTime : Time;
   END_VAR
   VAR_IN_OUT
      PressRam : "FB_CylinderCM";
      Door : "FB_CylinderCM";
      PartSlide : "FB_CylinderCM";
      Core : "FRK_Core";
      Unit : "FRK_Unit";
      Status : "ST_ModuleStatus";
      Part : "ST_PartContext";
      AlarmLog : "FRK_AlarmLog";
      Chart : "FB_GRAPH_PressDemoAuto";
   END_VAR
   VAR
      Seq { ExternalWritable := 'False'; S7_SetPoint := 'True'} : "FRK_SequenceCtx";
      Row1 { ExternalWritable := 'False'; S7_SetPoint := 'True'} : "FRK_SequenceRow";
      Row2 { ExternalWritable := 'False'; S7_SetPoint := 'True'} : "FRK_SequenceRow";
      Row3 { ExternalWritable := 'False'; S7_SetPoint := 'True'} : "FRK_SequenceRow";
      Row4 { ExternalWritable := 'False'; S7_SetPoint := 'True'} : "FRK_SequenceRow";
      Row5 { ExternalWritable := 'False'; S7_SetPoint := 'True'} : "FRK_SequenceRow";
      Row6 { ExternalWritable := 'False'; S7_SetPoint := 'True'} : "FRK_SequenceRow";
      Row7 { ExternalWritable := 'False'; S7_SetPoint := 'True'} : "FRK_SequenceRow";
      Row8 { ExternalWritable := 'False'; S7_SetPoint := 'True'} : "FRK_SequenceRow";
      Row9 { ExternalWritable := 'False'; S7_SetPoint := 'True'} : "FRK_SequenceRow";
      Row10 { ExternalWritable := 'False'; S7_SetPoint := 'True'} : "FRK_SequenceRow";
      Row11 { ExternalWritable := 'False'; S7_SetPoint := 'True'} : "FRK_SequenceRow";
      Row12 { ExternalWritable := 'False'; S7_SetPoint := 'True'} : "FRK_SequenceRow";
      Row13 { ExternalWritable := 'False'; S7_SetPoint := 'True'} : "FRK_SequenceRow";
      Row14 { ExternalWritable := 'False'; S7_SetPoint := 'True'} : "FRK_SequenceRow";
      Row15 { ExternalWritable := 'False'; S7_SetPoint := 'True'} : "FRK_SequenceRow";
      Row16 { ExternalWritable := 'False'; S7_SetPoint := 'True'} : "FRK_SequenceRow";
      At0 { ExternalAccessible := 'False'; ExternalVisible := 'False'; ExternalWritable := 'False'} : Bool;
      At100 { ExternalAccessible := 'False'; ExternalVisible := 'False'; ExternalWritable := 'False'} : Bool;
      At110 { ExternalAccessible := 'False'; ExternalVisible := 'False'; ExternalWritable := 'False'} : Bool;
      At130 { ExternalAccessible := 'False'; ExternalVisible := 'False'; ExternalWritable := 'False'} : Bool;
      At150 { ExternalAccessible := 'False'; ExternalVisible := 'False'; ExternalWritable := 'False'} : Bool;
      At170 { ExternalAccessible := 'False'; ExternalVisible := 'False'; ExternalWritable := 'False'} : Bool;
      At180 { ExternalAccessible := 'False'; ExternalVisible := 'False'; ExternalWritable := 'False'} : Bool;
      At185 { ExternalAccessible := 'False'; ExternalVisible := 'False'; ExternalWritable := 'False'} : Bool;
      At190 { ExternalAccessible := 'False'; ExternalVisible := 'False'; ExternalWritable := 'False'} : Bool;
      At200 { ExternalAccessible := 'False'; ExternalVisible := 'False'; ExternalWritable := 'False'} : Bool;
      At210 { ExternalAccessible := 'False'; ExternalVisible := 'False'; ExternalWritable := 'False'} : Bool;
      At215 { ExternalAccessible := 'False'; ExternalVisible := 'False'; ExternalWritable := 'False'} : Bool;
      At220 { ExternalAccessible := 'False'; ExternalVisible := 'False'; ExternalWritable := 'False'} : Bool;
      At230 { ExternalAccessible := 'False'; ExternalVisible := 'False'; ExternalWritable := 'False'} : Bool;
      At240 { ExternalAccessible := 'False'; ExternalVisible := 'False'; ExternalWritable := 'False'} : Bool;
      At999 { ExternalAccessible := 'False'; ExternalVisible := 'False'; ExternalWritable := 'False'} : Bool;
      Ready1 { ExternalAccessible := 'False'; ExternalVisible := 'False'; ExternalWritable := 'False'} : Bool;
      Ready2 { ExternalAccessible := 'False'; ExternalVisible := 'False'; ExternalWritable := 'False'} : Bool;
      Ready3 { ExternalAccessible := 'False'; ExternalVisible := 'False'; ExternalWritable := 'False'} : Bool;
      Ready4 { ExternalAccessible := 'False'; ExternalVisible := 'False'; ExternalWritable := 'False'} : Bool;
      Ready5 { ExternalAccessible := 'False'; ExternalVisible := 'False'; ExternalWritable := 'False'} : Bool;
      Advance { ExternalAccessible := 'False'; ExternalVisible := 'False'; ExternalWritable := 'False'} : Bool;
      Cycle { ExternalAccessible := 'False'; ExternalVisible := 'False'; ExternalWritable := 'False'; S7_SetPoint := 'True'} : "ST_PressDemoCycle";
      LoadPosition { ExternalAccessible := 'False'; ExternalVisible := 'False'; ExternalWritable := 'False'; S7_SetPoint := 'True'} : "FB_PressDemoLoadPosition";
      LoadDone { ExternalAccessible := 'False'; ExternalVisible := 'False'; ExternalWritable := 'False'} : Bool;
      LoadActive { ExternalAccessible := 'False'; ExternalVisible := 'False'; ExternalWritable := 'False'} : Bool;
      Branch1 { ExternalAccessible := 'False'; ExternalVisible := 'False'; ExternalWritable := 'False'; S7_SetPoint := 'True'} : "FRK_SequenceCtx";
      Branch2 { ExternalAccessible := 'False'; ExternalVisible := 'False'; ExternalWritable := 'False'; S7_SetPoint := 'True'} : "FRK_SequenceCtx";
      Row17 { ExternalWritable := 'False'; S7_SetPoint := 'True'} : "FRK_SequenceRow";
      Row18 { ExternalWritable := 'False'; S7_SetPoint := 'True'} : "FRK_SequenceRow";
      Row19 { ExternalWritable := 'False'; S7_SetPoint := 'True'} : "FRK_SequenceRow";
   END_VAR
BEGIN

   "FRK_SeqBegin"(Run := #Run,
                  Reset := #Reset,
                  OwnerIndex := #OwnerIndex,
                  ChainIndex := 1,
                  BranchIndex := 0,
                  Delta := #Delta,
                  Seq := #Seq);
   "FRK_SeqStart"(Seq := #Seq,
                  StartPulse := #StartPulse);
   "F_PressDemoReset"(Seq := #Seq,
                      Cycle := #Cycle);
   "FRK_SeqBegin"(Run := #Run,
                  Reset := #Reset,
                  OwnerIndex := #OwnerIndex,
                  ChainIndex := 1,
                  BranchIndex := 1,
                  Delta := #Delta,
                  Seq := #Branch1);
   "FRK_SeqBegin"(Run := #Run,
                  Reset := #Reset,
                  OwnerIndex := #OwnerIndex,
                  ChainIndex := 1,
                  BranchIndex := 2,
                  Delta := #Delta,
                  Seq := #Branch2);
   #LoadActive := "FRK_SeqSubActive"(Seq := #Branch1, Run := #Run, StepNo := 240);
   #LoadDone := "F_PressDemoLoadPosition"(Target := #LoadPosition, Run := #LoadActive, Reset := #Seq.Restart, OwnerIndex := #OwnerIndex, Delta := #Delta, PressRam := #PressRam, Door := #Door, PartSlide := #PartSlide);
   "F_CylinderSequenceLease"(Seq := #Seq,
                             Target := #PressRam);
   "F_CylinderSequenceLease"(Seq := #Seq,
                             Target := #Door);
   "F_CylinderSequenceLease"(Seq := #Seq,
                             Target := #PartSlide);
   "F_CylinderSequenceLease"(Seq := #Branch1,
                             Target := #PressRam);
   "F_CylinderSequenceLease"(Seq := #Branch1,
                             Target := #Door);
   "F_CylinderSequenceLease"(Seq := #Branch1,
                             Target := #PartSlide);
   "F_CylinderSequenceLease"(Seq := #Branch2,
                             Target := #PressRam);
   "F_CylinderSequenceLease"(Seq := #Branch2,
                             Target := #Door);
   "F_CylinderSequenceLease"(Seq := #Branch2,
                             Target := #PartSlide);
   #Chart(Run := #Run,
          Reset := #Reset,
          OwnerIndex := #OwnerIndex,
          Delta := #Delta,
          TransferSettleTime := #TransferSettleTime,
          PartQuality := #PartQuality,
          RequireTwoHandStart := #RequireTwoHandStart,
          SourcePath := #SourcePath,
          PartPresent := #PartPresent,
          AirPressureOk := #AirPressureOk,
          TwoHandHeld := #TwoHandHeld,
          StartPulse := #StartPulse,
          PressSettleTime := #PressSettleTime,
          PressRam := #PressRam,
          Door := #Door,
          PartSlide := #PartSlide,
          HostCore := #Core,
          HostUnit := #Unit,
          HostStatus := #Status,
          HostPart := #Part,
          HostAlarmLog := #AlarmLog,
          Seq := #Seq,
          Row1 := #Row1,
          Row2 := #Row2,
          Row3 := #Row3,
          Row4 := #Row4,
          Row5 := #Row5,
          Row6 := #Row6,
          Row7 := #Row7,
          Row8 := #Row8,
          Row9 := #Row9,
          Row10 := #Row10,
          Row11 := #Row11,
          Row12 := #Row12,
          Row13 := #Row13,
          Row14 := #Row14,
          Row15 := #Row15,
          Row16 := #Row16,
          Ready1 := #Ready1,
          Ready2 := #Ready2,
          Ready3 := #Ready3,
          Ready4 := #Ready4,
          Ready5 := #Ready5,
          Cycle := #Cycle,
          LoadDone := #LoadDone,
          Branch1 := #Branch1,
          Branch2 := #Branch2,
          Row17 := #Row17,
          Row18 := #Row18,
          Row19 := #Row19,
          INIT_SQ := #Seq.Restart,
          OFF_SQ := NOT #Seq.Running);
   "FRK_SeqSubStatus"(Seq := #Branch1,
                      Child := #LoadPosition.Seq);
   "FRK_SeqOwnerStatus"(Seq := #Branch1,
                        Core := #Core,
                        Status := #Status);
   "FRK_SeqOwnerStatus"(Seq := #Branch2,
                        Core := #Core,
                        Status := #Status);
   "FRK_SeqOwnerStatus"(Seq := #Seq,
                        Core := #Core,
                        Status := #Status);
   "F_CylinderSequenceLease"(Seq := #Seq,
                             Target := #PressRam);
   "F_CylinderSequenceLease"(Seq := #Seq,
                             Target := #Door);
   "F_CylinderSequenceLease"(Seq := #Seq,
                             Target := #PartSlide);
   "F_CylinderSequenceLease"(Seq := #Branch1,
                             Target := #PressRam);
   "F_CylinderSequenceLease"(Seq := #Branch1,
                             Target := #Door);
   "F_CylinderSequenceLease"(Seq := #Branch1,
                             Target := #PartSlide);
   "F_CylinderSequenceLease"(Seq := #Branch2,
                             Target := #PressRam);
   "F_CylinderSequenceLease"(Seq := #Branch2,
                             Target := #Door);
   "F_CylinderSequenceLease"(Seq := #Branch2,
                             Target := #PartSlide);
END_FUNCTION_BLOCK

